(* IEC 61131-3 sources: daoli-st-library/DL_Device (part 15) *)

(* ---- FB_DL_CaseErectFaultSeq.st ---- *)
(*==============================================================================
 * 组件名称 (Component)  : FB_DL_CaseErectFaultSeq
 * 所属子库 (Sublibrary) : DL_Device
 * 当前版本 (Version)    : 1.0.0
 * 兼容性 (Platform)     : CODESYS 3.5+ / TwinCAT 3 / 汇川 InoProShop / 施耐德 Machine Expert
 *                         仅依赖 Standard.library（TON / R_TRIG），零厂商私有库
 * 功能描述 (Function)   : 开箱成型失败重试与吸盘堵塞诊断。bStartCmd 沿启动
 *                         成型吸持：bSuctionCmd 置位等待真空达 fVacOkLevel
 *                         （tonSeek 窗）；达压 → bPickDone 单拍并保持吸持监视
 *                         （中途掉压判 eVacDrop）；超时 → 吹气清理（bBlowOffCmd
 *                         in eRetryPause tRetryPause）后重试，超 nMaxRetry 次
 *                         归因收口：全程真空峰值 <= fVacFloor → eVacClog（吸盘
 *                         堵塞/无真空），曾达压后掉 → eVacDrop，部分真空但
 *                         不足 → eVacTimeout。三成因独立分码（R190 归因唯一）。
 * 来源标签 (Origin)     : ROADMAP 在册空勾 P2（R13 新增行）；判据思想复用既有
 *                         VacuumEjector 件（真空等级判据语义域借鉴），实现与
 *                         码位独立 clean-room，IEC 61131-3 标准语义的道莅防御性实现
 * 边界语义 (Boundary)   : ① 三段 TON 一相一实例（R275）：tonSeek/tonPause/
 *                         tonDrop 各自独立，禁跨相复用；
 *                         ② 归因锁存：故障相按锁存回放，不按当下真空重推断（R28）；
 *                         ③ 重试计数只在收口沿或复位沿清（bStop 中止保留计数，
 *                         作用域在此声明——中止视为本轮未完，重试额度保留）；
 *                         ④ 组态闸：真空等级/地板值/时间/次数全引脚覆盖（R151）。
 * 输出语义 (Fallback)   : 【R191】bEnable = FALSE → 全输出强制 FALSE（吸持是
 *                         执行器指令，失能必须收敛）；eFault 相 → bSuctionCmd
 *                         强制 FALSE（故障先断气源），bError = TRUE。
 * 码位     (Codes)      : 按 R297 范式零 16# 码位硬编码；错误出口 BOOL+ENUM(eCause)，
 *                         码位待主控收口统一派号。
 * 红线自检 (Redline)    : 7 项红线已自检：R1 零全局 ✓｜R2 零物理地址 ✓｜R3 纯 IEC ✓
 *                         R4 组态闸全引脚/容差比较 ✓｜R5 双语同行注释 ✓
 *                         R6 CASE 带 ELSE 兜底迁 eFault ✓
 *                         R7 三 TON + 两 R_TRIG 段 0 无条件刷新，各实例单用途 ✓
 * 验收向量 (Acceptance) : V1 首次达压 → bPickDone 单拍 TRUE，nRetryCnt=0；
 *                         V2 达压后掉压 → eFault，eCause=eVacDrop；
 *                         V3 三次超时且真空峰值恒为地板值 → eCause=eVacClog；
 *                         V4 三次超时峰值 0.5·fVacOkLevel → eCause=eVacTimeout；
 *                         V5 重试期 bBlowOffCmd 电平 TRUE（暂停相内）。
 * 修订历史 (Revision)   : 2026-11-20  v1.0.0  R49 首版（批 2 · 序号 10）
 *==============================================================================*)
TYPE E_DL_CefState :
(
    eIdle       := 0,                        (* 待启动 / Idle *)
    eErect      := 10,                       (* 吸持建立中（真空达压窗） / Erecting, vacuum seek *)
    eHold       := 20,                       (* 吸持保持监视（掉压判据） / Holding, drop watch *)
    eRetryPause := 30,                       (* 吹气清理暂停（重试间隔） / Blow-off pause *)
    eFault      := 90                        (* 故障锁存相 / Fault latched phase *)
);
END_TYPE

TYPE E_DL_CefCause :
(
    eNone        := 0,                       (* 无故障成因 / No cause *)
    eVacClog     := 1,                       (* 吸盘堵塞：全程真空不高于地板值 / Suction clog: vacuum never above floor *)
    eVacDrop     := 2,                       (* 中途掉压：曾达压后失压 / Vacuum drop after reaching level *)
    eVacTimeout  := 3,                       (* 达压超时：部分真空但始终不足 / Vacuum seek timeout, partial only *)
    eCfgIllegal  := 4,                       (* 组态非法 / Illegal config *)
    ePhaseBad    := 5                        (* 非法相位兜底 / Illegal phase fallback *)
);
END_TYPE

FUNCTION_BLOCK FB_DL_CaseErectFaultSeq
VAR_INPUT
    bVacOkLvl   : BOOL := FALSE;             (* 真空达压电平（真空开关或比较器输出直连）[-] / Vacuum-ok level input *)
    fVacReading : LREAL := 0.0;              (* 真空读数（归因诊断用）[kPa] / Vacuum reading for diagnosis *)
    fVacOkLevel : LREAL := 60.0;             (* 达压等级阈值，域 > 0.0 [kPa] / Vacuum ok threshold *)
    fVacFloor   : LREAL := 5.0;              (* 地板值：峰值不高于此判堵塞，域 >= 0.0 且 < fVacOkLevel [kPa] / Vacuum floor for clog verdict *)
    tVacSeek    : TIME := T#3S;              (* 达压窗保持时长，域 > T#0S [ms] / Vacuum seek window *)
    tRetryPause : TIME := T#1S;              (* 吹气清理暂停保持时长，域 > T#0S [ms] / Retry pause hold *)
    nMaxRetry   : INT := 3;                  (* 最大重试次数，域 0..20 [次] / Max retry count *)
    bStartCmd   : BOOL := FALSE;             (* 成型启动命令，上升沿发起 / Start command edge *)
    bStop       : BOOL := FALSE;              (* 中止命令，电平 TRUE 立即断吸回 eIdle（保留重试计数，见边界③） / Stop level, keeps retry count *)
    bEnable     : BOOL := TRUE;              (* 使能，FALSE 全输出强制收敛 [-] / Enable *)
    bReset      : BOOL := FALSE;              (* 复位命令，上升沿清故障锁存与全部状态 [-] / Reset command *)
END_VAR
VAR_OUTPUT
    bSuctionCmd : BOOL;                      (* 吸盘吸持命令输出 [-] / Suction command output *)
    bBlowOffCmd : BOOL;                      (* 吹气清理命令输出（重试暂停相电平）[-] / Blow-off command output *)
    bPickDone   : BOOL;                      (* 本轮吸持达压完成单拍位 [-] / Pick-done single-scan pulse *)
    nRetryCnt   : INT;                       (* 本轮已用重试次数 [次] / Retry count this round *)
    nAttemptCnt : INT;                       (* 本轮尝试总次数（含首次）[次] / Attempt count this round *)
    eState      : E_DL_CefState;             (* 状态出口 / State outlet *)
    eCause      : E_DL_CefCause;             (* 故障成因出口（R190 三成因独立分码） / Fault cause outlet *)
    bError      : BOOL;                       (* 故障锁存标志 [-] / Fault latch flag *)
END_VAR
VAR
    _eState   : E_DL_CefState := E_DL_CefState.eIdle;     (* 内部相位（CASE 唯一写入目标） / Internal phase *)
    _eCause   : E_DL_CefCause := E_DL_CefCause.eNone;     (* 故障成因锁存量 / Latched cause *)
    tonSeek   : TON;                         (* 达压窗计时（eErect 相专用），段 0 无条件调用 / Seek timer, phase-specific *)
    tonPause  : TON;                         (* 吹气暂停计时（eRetryPause 相专用），段 0 无条件调用 / Pause timer, phase-specific *)
    tonDrop   : TON;                         (* 掉压确认计时（eHold 相专用），段 0 无条件调用 / Drop confirm timer, phase-specific *)
    rtStart   : R_TRIG;                      (* 启动沿实例，段 0 无条件调用 / Start edge instance *)
    rtReset   : R_TRIG;                      (* 复位沿实例，段 0 无条件调用 / Reset edge instance *)
    _nRetry   : INT;                         (* 重试计数锁存 [次] / Retry count latch *)
    _nAttempt : INT;                         (* 尝试计数锁存 [次] / Attempt count latch *)
    _fVacMax  : LREAL;                       (* 本轮真空峰值锁存（归因判据源）[kPa] / Vacuum peak latch *)
    _bReached : BOOL;                        (* 本轮曾达压位（掉压归因判据）[-] / Reached-ok latch this round *)
    _bFault   : BOOL;                        (* 故障锁存位 / Latched fault bit *)
    _bCfgBad  : BOOL;                        (* 组态非法当拍量 / Illegal config this scan *)
END_VAR

(* —— 段 0：当拍判据派生 + 实例无条件刷新（R228A，三 TON 各自独立 IN 派生） —— *)
_bCfgBad := (fVacOkLevel <= 0.0) OR (fVacFloor < 0.0) OR (fVacFloor >= fVacOkLevel)   (* 组态闸：等级/地板域及序关系（R151 全引脚覆盖） / Config gate *)
            OR (tVacSeek <= T#0S) OR (tRetryPause <= T#0S) OR (nMaxRetry < 0) OR (nMaxRetry > 20);
rtStart(CLK := bStartCmd);                   (* 启动沿每拍必调 / Start edge every scan *)
rtReset(CLK := bReset);                      (* 复位沿每拍必调 / Reset edge every scan *)
tonSeek(IN := _eState = E_DL_CefState.eErect, PT := tVacSeek);        (* 达压窗随相位派生 / Seek timer phase-derived *)
tonPause(IN := _eState = E_DL_CefState.eRetryPause, PT := tRetryPause);   (* 暂停计时随相位派生 / Pause timer phase-derived *)
tonDrop(IN := _eState = E_DL_CefState.eHold AND NOT bVacOkLvl, PT := tRetryPause);   (* 掉压确认随相位派生（PT 复用暂停时长作为失压容忍窗，语义声明） / Drop confirm timer *)

(* —— 段 1：单拍量预清零（R107） —— *)
bPickDone := FALSE;                          (* 达压完成单拍位预清，唯一分支置位 / Pick pulse preset *)

(* —— 段 2：复位沿处理（作用域：清故障 + 清成因 + 清计数 + 清峰值 + 迁 eIdle，R283 逐项声明） —— *)
IF rtReset.Q THEN
    _bFault := FALSE;                        (* 清故障锁存 / Clear fault *)
    _eCause := E_DL_CefCause.eNone;          (* 清成因 / Clear cause *)
    _nRetry := 0;                            (* 清重试计数 / Clear retry count *)
    _nAttempt := 0;                          (* 清尝试计数 / Clear attempt count *)
    _fVacMax := 0.0;                         (* 清真空峰值 / Clear vacuum peak *)
    _bReached := FALSE;                      (* 清曾达压位 / Clear reached latch *)
    _eState := E_DL_CefState.eIdle;          (* 迁待启动相 / Back to idle *)
END_IF

(* —— 段 3：组态闸故障锁存（R45 配对；锁存至复位沿，R189） —— *)
IF _bCfgBad AND NOT _bFault THEN
    _bFault := TRUE;                         (* 锁存故障位 / Latch fault *)
    _eCause := E_DL_CefCause.eCfgIllegal;    (* 成因：组态非法 / Cause: illegal config *)
    _eState := E_DL_CefState.eFault;         (* 同步迁故障相 / Migrate to fault *)
END_IF

(* —— 段 4：CASE 主状态机（ELSE 兜底迁 eFault，红线 6） —— *)
CASE _eState OF
    E_DL_CefState.eIdle:                     (* 待启动相 / Idle *)
        IF rtStart.Q AND bEnable AND NOT _bFault THEN
            _nAttempt := _nAttempt + 1;      (* 尝试计数递增 / Attempt count advance *)
            _fVacMax := 0.0;                 (* 本轮峰值清零 / Clear round peak *)
            _bReached := FALSE;              (* 本轮曾达压清零 / Clear reached latch *)
            _eState := E_DL_CefState.eErect; (* 进入吸持建立 / Enter erect *)
        END_IF
    E_DL_CefState.eErect:                    (* 吸持建立相 / Erect *)
        IF NOT bEnable OR bStop THEN         (* 失能/中止：断吸回待机（重试计数保留，边界③声明） / Disable or stop *)
            _eState := E_DL_CefState.eIdle;  (* 回待机 / Back to idle *)
        ELSIF bVacOkLvl THEN
            _bReached := TRUE;               (* 曾达压置位 / Reached latch *)
            bPickDone := TRUE;               (* 达压完成单拍脉冲 / Pick-done pulse *)
            _eState := E_DL_CefState.eHold;  (* 进入保持监视 / Enter hold *)
        ELSE
            IF fVacReading > _fVacMax THEN
                _fVacMax := fVacReading;     (* 真空峰值跟踪（NaN 参与比较恒 FALSE，不污染峰值） / Vacuum peak tracking, NaN-safe *)
            END_IF
            IF tonSeek.Q THEN
                _nRetry := _nRetry + 1;      (* 超时计一次重试 / Retry count advance *)
                IF _nRetry > nMaxRetry THEN
                    IF _bReached THEN
                        _eCause := E_DL_CefCause.eVacDrop;      (* 曾达压后失压归因（独立分码，R190） / Drop cause *)
                    ELSIF _fVacMax <= fVacFloor THEN
                        _eCause := E_DL_CefCause.eVacClog;      (* 峰值不高于地板：吸盘堵塞归因 / Clog cause *)
                    ELSE
                        _eCause := E_DL_CefCause.eVacTimeout;   (* 部分真空但不足：超时归因 / Timeout cause *)
                    END_IF
                    _bFault := TRUE;         (* 重试耗尽故障锁存（R45 配对） / Retry exhausted fault *)
                    _eState := E_DL_CefState.eFault;   (* 同步迁故障相 / Migrate to fault *)
                ELSE
                    _eState := E_DL_CefState.eRetryPause;   (* 未耗尽：吹气清理后重试 / Enter retry pause *)
                END_IF
            END_IF
        END_IF
    E_DL_CefState.eHold:                     (* 吸持保持相 / Hold *)
        IF NOT bEnable OR bStop THEN
            _eState := E_DL_CefState.eIdle;  (* 失能/中止回待机 / Back to idle *)
        ELSIF bVacOkLvl THEN
            ;                                (* 吸持正常，无动作 / Holding normal *)
        ELSIF tonDrop.Q THEN                 (* 失压持续到容忍窗 / Drop held to tolerance *)
            _eCause := E_DL_CefCause.eVacDrop;   (* 中途掉压归因（独立分码，R190） / Drop cause *)
            _bFault := TRUE;                 (* 故障锁存（R45 配对） / Latch fault *)
            _eState := E_DL_CefState.eFault; (* 同步迁故障相 / Migrate to fault *)
        END_IF
    E_DL_CefState.eRetryPause:               (* 吹气清理暂停相 / Retry pause *)
        IF NOT bEnable OR bStop THEN
            _eState := E_DL_CefState.eIdle;  (* 失能/中止回待机 / Back to idle *)
        ELSIF tonPause.Q THEN
            _nAttempt := _nAttempt + 1;      (* 新尝试计数 / Attempt count advance *)
            _eState := E_DL_CefState.eErect; (* 重新吸持建立 / Re-enter erect *)
        END_IF
    E_DL_CefState.eFault:                    (* 故障相：先断气源，仅复位沿出 / Fault: suction cut *)
        ;                                    (* 锁存回放（R28） / Replay from latch *)
    ELSE                                     (* 非法相位兜底迁安全态 / Illegal phase fallback *)
        _eState := E_DL_CefState.eFault;     (* 迁故障相 / To fault *)
        _bFault := TRUE;                     (* 同步锁存 / Latch *)
        _eCause := E_DL_CefCause.ePhaseBad;  (* 成因：非法相位 / Cause: illegal phase *)
END_CASE

(* —— 段 5：出口映射（双门控：失能收敛 + 故障断气源，R191/R285 全路径赋值） —— *)
IF (NOT bEnable) OR _bFault OR (_eState = E_DL_CefState.eIdle) THEN
    bSuctionCmd := FALSE;                    (* 失能/故障/待机：吸持强制收敛 / Suction forced off *)
    bBlowOffCmd := FALSE;                    (* 吹气强制收敛 / Blow-off forced off *)
ELSIF _eState = E_DL_CefState.eErect OR _eState = E_DL_CefState.eHold THEN
    bSuctionCmd := TRUE;                     (* 建立/保持相：吸持命令电平 / Suction on *)
    bBlowOffCmd := FALSE;                    (* 吹气关闭 / Blow-off off *)
ELSIF _eState = E_DL_CefState.eRetryPause THEN
    bSuctionCmd := FALSE;                    (* 暂停相断吸 / Suction off *)
    bBlowOffCmd := TRUE;                     (* 吹气清理电平 / Blow-off on *)
ELSE
    bSuctionCmd := FALSE;                    (* 兜底收敛 / Fallback off *)
    bBlowOffCmd := FALSE;                    (* 兜底收敛 / Fallback off *)
END_IF
nRetryCnt := _nRetry;                        (* 重试计数镜像 / Retry count mirror *)
nAttemptCnt := _nAttempt;                    (* 尝试计数镜像 / Attempt count mirror *)
bError := _bFault;                           (* 故障标志镜像 / Fault flag mirror *)
eState := _eState;                           (* 状态出口 / State outlet *)
eCause := _eCause;                           (* 成因出口 / Cause outlet *)
END_FUNCTION_BLOCK

(* ---- FB_DL_CaseSealTapeMonitor.st ---- *)
(*
  FB_DL_CaseSealTapeMonitor  —  封箱胶带缺料/断带监视 / Case sealing tape run-out and break monitor
  分类 Category : DL_Device
  码位 Code     : 16#03_2_0A
  版本 Version  : 1.0.0
  溯源 Source   : ISA-18.2 报警管理语义借鉴 · clean-room 实现，仅借分类/参数域/命名，未复制源码
  功能 Function : 1) 张力 + 光电双判据封箱胶带状态监视（复用 FB_DL_SignalDebounce 去抖）；
                  2) 节拍使能时连续 N 拍「无张力 + 光电同态」才判断带（防单拍尖峰）；
                  3) 缺料与断带独立码值（FB33-3 归因唯一），解除需补料确认 + 复位沿。
  边界 Boundary : ① 节拍使能时连续 N 拍无张力 + 光电同态才判断带（防单拍尖峰）；
                  ② 张力传感器无效冻结判定并置码；
                  ③ 缺料（低张力 + 光电无带）与断带（运动中张力突失）独立码值；
                  ④ 报警解除需补料确认 + 复位沿（双条件可达）；
                  ⑤ 输出三行同向：缺料 → 断带 → 去抖状态。
  依赖 Depends  : FB_DL_SignalDebounce × 2（张力低 / 光电无带去抖，每拍无条件调用）

  码表 Error codes（本件子码步进 16#10，避让邻件码位）:
    16#0002_030A 故障级：组态非法（确认拍数 < 1 / 去抖时长 < 0）
    16#0002_031A 故障级：断带（运动中张力突失 + 光电同态确认，锁存需补料 + 复位沿）
    16#0002_032A 信息级：缺料（低张力 + 光电无带，提示级）/ 张力无效判定冻结（不置 bError）
*)

TYPE E_DL_CstPhase :
(
    eIdle  := 0,  // 空闲 / Idle
    eWatch := 10, // 胶带状态监视 / Tape watching
    eBreak := 20, // 断带锁存 / Tape break latched
    eFault := 90  // 组态故障锁定 / Configuration fault locked
);
END_TYPE

FUNCTION_BLOCK FB_DL_CaseSealTapeMonitor
VAR_INPUT
    bEnable       : BOOL;                           // 总使能，FALSE 回空闲 / Master enable
    bCycleEn      : BOOL;                           // 封箱节拍使能（运动中判定窗口）/ Sealing cycle enable
    bReset        : BOOL;                           // 复位，上升沿清组态故障 / Reset, clears fault
    fTensionN     : REAL;                           // 胶带张力 [N] / Tape tension [N]
    bPhotoSensor  : BOOL;                           // 光电传感（TRUE = 有带）/ Photo sensor, TRUE = tape present
    fTensionLoN   : REAL := 2.0;                    // 张力下限 [N]（低于判无张力）/ Tension low limit [N]
    uBreakConfirm : UINT := 5;                      // 断带确认拍数 [拍] / Break confirm scans
    tDebounce     : TIME := T#100MS;                // 信号去抖时长 [ms] / Signal debounce time
    bTapeRefeed   : BOOL;                           // 补料确认（解除条件之一）/ Tape refeed confirmed
    fEps          : REAL := 1.0E-6;                 // 浮点判零容差 [1] / Floating zero tolerance
END_VAR
VAR_OUTPUT
    bTapeMissing  : BOOL;                           // 缺料标志（提示级）/ Tape missing flag, info level
    bTapeBreak    : BOOL;                           // 断带标志（锁存）/ Tape break flag, latched
    bDebouncing   : BOOL;                           // 去抖进行中标志 / Debouncing flag
    bError        : BOOL;                           // 故障标志，与故障级码配对 / Fault flag
    uErrorId      : UDINT;                          // 事件码，0 = 无事件 / Event code
    eStateOut     : E_DL_CstPhase;                  // 状态机当前态，段尾单点映射 / Phase mapped at tail
END_VAR
VAR
    _eState       : E_DL_CstPhase := E_DL_CstPhase.eIdle;  // 内部状态 / Internal state
    fbDebTension  : FB_DL_SignalDebounce;           // 张力低去抖实例（无条件调用）/ Tension-low debounce
    fbDebPhoto    : FB_DL_SignalDebounce;           // 光电无带去抖实例（无条件调用）/ Photo-no-tape debounce
    rtrReset      : R_TRIG;                         // 复位沿 / Reset edge
    bCfgOk        : BOOL;                           // 组态合法标志 / Configuration valid
    bTensionOk    : BOOL;                           // 张力本拍有效 / Tension valid this scan
    bNoTension    : BOOL;                           // 无张力（去抖后）/ No tension, debounced
    bNoPhoto      : BOOL;                           // 光电无带（去抖后）/ No tape by photo, debounced
    bBreakCond    : BOOL;                           // 断带条件（无张力 + 光电同态）/ Break condition
    uBreakCnt     : UINT;                           // 断带确认计数 [拍] / Break confirm counter
    uFault        : UDINT;                          // 锁存故障码 / Latched fault code
    uInfo         : UDINT;                          // 信息级码 / Information code
END_VAR

(* === 段 0 · 实例刷新 === *)
rtrReset(CLK := bReset);                          // 每拍刷新复位沿

(* === 段 1 · 组态闸 === *)
bCfgOk := (uBreakConfirm >= UINT#1)               // 确认拍数下限
          AND (TIME_TO_REAL(tDebounce) >= 0.0)    // 去抖时长非负
          AND (fTensionLoN >= 0.0)                // 张力下限非负域
          AND (fTensionLoN = fTensionLoN);        // NaN 自反
IF NOT bCfgOk THEN
    uFault := 16#0002_030A;                       // 故障级：组态非法
END_IF
IF rtrReset.Q AND bCfgOk THEN
    uFault := 16#0000;                            // 复位沿清组态锁存（解除路径可达）
END_IF
uInfo := 16#0000;                                 // 信息码每拍清零
bTensionOk := (fTensionN = fTensionN) AND (fTensionN >= 0.0) AND (fTensionN < 1.0E30);  // 张力 NaN 自反 + 非负域

(* === 段 2 · 去抖实例（无条件调用）与双判据合成 === *)
fbDebTension(bRawInput := bTensionOk AND (fTensionN < fTensionLoN),   // 原始判据：张力低于下限
             tRiseDelay := tDebounce,             // 上升去抖
             tFallDelay := tDebounce,             // 下降去抖
             bEnable := bEnable AND bCfgOk,       // 使能透传
             bReset := rtrReset.Q);               // 复位沿透传
fbDebPhoto(bRawInput := (NOT bPhotoSensor),       // 原始判据：光电无带
           tRiseDelay := tDebounce,               // 上升去抖
           tFallDelay := tDebounce,               // 下降去抖
           bEnable := bEnable AND bCfgOk,         // 使能透传
           bReset := rtrReset.Q);                 // 复位沿透传
bNoTension := fbDebTension.bStable;               // 无张力（去抖后）
bNoPhoto := fbDebPhoto.bStable;                   // 光电无带（去抖后）
bDebouncing := fbDebTension.bFiltering OR fbDebPhoto.bFiltering;   // 去抖进行中
bBreakCond := bCycleEn AND bTensionOk AND bNoTension AND bNoPhoto;  // 节拍使能 + 无张力 + 光电同态
bTapeMissing := (NOT bCycleEn) AND bTensionOk AND bNoTension AND bNoPhoto;   // 非节拍缺料（提示级）
IF NOT bTensionOk THEN
    uInfo := 16#0002_032A;                        // 信息级：张力无效判定冻结
    uBreakCnt := UINT#0;                          // 无效拍计数归零（禁污染确认）
END_IF

(* === 段 3 · 断带确认计数（连续 N 拍防单拍尖峰）=== *)
IF bBreakCond THEN
    uBreakCnt := uBreakCnt + UINT#1;              // 断带条件确认计数
    IF uBreakCnt >= uBreakConfirm THEN
        uFault := 16#0002_031A;                   // 故障级：断带锁存（需补料 + 复位沿）
    END_IF
ELSE
    uBreakCnt := UINT#0;                          // 条件消失计数归零
END_IF
bTapeBreak := (uFault = 16#0002_031A);            // 断带出口（锁存态映射）

(* === 段 4 · 主状态机（ENUM + CASE，含 ELSE 兜底）=== *)
CASE _eState OF
E_DL_CstPhase.eIdle :
    IF uFault <> 16#0000 THEN
        _eState := E_DL_CstPhase.eFault;          // 故障优先
    ELSIF bEnable AND bCfgOk THEN
        _eState := E_DL_CstPhase.eWatch;          // 进监视相
    END_IF

E_DL_CstPhase.eWatch :
    IF uFault <> 16#0000 THEN
        _eState := E_DL_CstPhase.eBreak;          // 断带锁存转断带相
    ELSIF (NOT bEnable) OR (NOT bCfgOk) THEN
        _eState := E_DL_CstPhase.eIdle;           // 失能回空闲
    END_IF

E_DL_CstPhase.eBreak :
    (* 解除条件：补料确认 + 复位沿（双条件齐备，路径可达） *)
    IF bTapeRefeed AND rtrReset.Q THEN
        uFault := 16#0000;                        // 复位沿清断带锁存
        uBreakCnt := UINT#0;                      // 确认计数复位
        _eState := E_DL_CstPhase.eWatch;          // 回监视相
    END_IF

E_DL_CstPhase.eFault :
    IF uFault = 16#0000 THEN
        _eState := E_DL_CstPhase.eIdle;           // 解锁回空闲
    END_IF

ELSE
    _eState := E_DL_CstPhase.eFault;              // 非法状态拦截
    uFault := 16#0002_030A;                       // 故障级：相 ID 越界复用组态码段
END_CASE

(* === 段 5 · 输出映射（缺料与断带归因唯一：独立码值独立出口）=== *)
IF NOT bTapeBreak THEN
    bTapeMissing := bTapeMissing AND bTensionOk AND bCfgOk;   // 非断带时缺料提示有效
END_IF
bError := (uFault <> 16#0000);                    // 故障标志仅由故障级码置位（R45 配对）
IF bError THEN
    uErrorId := uFault;                           // 故障级优先上报
ELSE
    uErrorId := uInfo;                            // 否则上报信息级码
END_IF
eStateOut := _eState;                             // 输出枚举段尾单点映射（N2 规则）
END_FUNCTION_BLOCK

(* ---- FB_DL_CellFeederVacuum.st ---- *)
(*
  FB_DL_CellFeederVacuum  —  电芯真空上料吸盘（真空窗 + 泄漏率判据 + 掉料重试） / Cell feeder vacuum cup with vacuum window, leakage-rate verdict and drop retry
  分类 Category : DL_Device
  版本 Version  : 1.0.0
  来源 Source   : t1-5-tcopen — 电芯上料吸盘执行器族深化
  溯源 Origin   : 道莅 clean-room 实现；真空窗确认 + 泄漏率判据 + 有限次重试为公开真空吸取工艺逻辑，未复制任何源码行
  功能 Function : 1) 三段顺控：eVac 抽真空（|fVacKpa - fVacTargetKpa| <= fVacTolKpa 达窗）→
                  eLeak 泄漏率测试窗（tLeak 内 fLeakKpaPerS <= fLeakMaxKpaPerS 且 bPartOn 在位）→
                  eDone；2) 掉料重试：泄漏/在位判据失败或 bPartOn 丢失 → eRetry 重抽，
                  重试计数 nRetry 达 nRetryMax 即故障（计数饱和于 nRetryMax）；
                  3) 抽真空超时、测试窗超时各自归因；
                  4) 故障级单码 052D / 信息级 0433 = 吸取确认完成沿。
  接口 Interface: 输入真空度/泄漏率/在位/三个时间量/重试上限；输出状态 + 吸盘指令 + 码
  边界 Boundary : ① 组态闸：fVacTargetKpa <= 0.0、fVacTolKpa <= 0.0、fLeakMaxKpaPerS <= 0.0、
                  tVacTmo/tLeak/tRetry <= T#0S、nRetryMax = 0 → 052D 锁存；
                  ② 真空度/泄漏率非有限（NaN 自反 + Inf 差值自减）→ 052D 锁存，吸盘保持指令撤销；
                  ③ 重试计数为 UINT，递增前先判饱和（不越界）；④ 三 TON + R_TRIG 段 0 无条件调用；
                  ⑤ 故障相迁出唯一路径 = bReset 上升沿（同时清重试计数）；
                  ⑥ 零全局耦合：无 GVL / VAR_EXTERNAL / %I %Q %M 直接地址。
  依赖 Depends  : Standard.library（TON / R_TRIG）
  码表 Error codes（Device 分段见下，故障窗口 052D / 信息窗口 0433）:
    16#0003_052D 故障级：真空上料故障总码（组态非法 / 抽真空超时 / 泄漏率超限且重试耗尽 / 输入非有限），
                 锁存至 bReset 上升沿；归因见 eCause，不新增码位（派单硬约束单码）
    16#0003_0433 信息级：吸取确认完成沿（进 eDone 单拍）
    分段理由：段 0003 故障带 03A0~03FF 于 R42 用尽，启用 05xx 副带续编，避开 0590~0599 判错位段。
  修订历史 Revision :
    2026-11-19  v1.0.0  R43 首版（批次 4 · 序号 17）
*)

TYPE E_DL_CfvState :
(
    eIdle   := 0,     // 未使能：吸盘指令撤销 / Idle, suction withdrawn
    eVac    := 10,    // 抽真空中 / Evacuating
    eLeak   := 20,    // 泄漏率测试窗 / Leakage test window
    eRetry  := 30,    // 掉料重试重抽中 / Retry re-evacuation
    eDone   := 50,    // 吸取完成 / Pick done
    eFault  := 90     // 故障锁存相 / Fault latched phase
);
END_TYPE

TYPE E_DL_CfvCause :
(
    eNone       := 0, // 无故障成因 / No cause
    eCfgIllegal := 1, // 组态非法 / Illegal configuration
    eVacTmo     := 2, // 抽真空超时 / Evacuation timeout
    eLeakHigh   := 3, // 泄漏率超限且重试耗尽 / Leakage high after retries
    eRetryOut   := 4, // 重试次数耗尽 / Retry exhausted
    eNonFinite  := 5  // 输入非有限 / Non-finite input
);
END_TYPE

FUNCTION_BLOCK FB_DL_CellFeederVacuum
VAR_INPUT
    fVacKpa        : REAL := 0.0;      // 吸盘真空度 [kPa]，正压差量纲 / Cup vacuum level
    fVacTargetKpa  : REAL := 60.0;     // 目标真空度 [kPa]，域 > 0 / Target vacuum level
    fVacTolKpa     : REAL := 3.0;      // 真空度容差 [kPa]，域 > 0 / Vacuum tolerance
    fLeakKpaPerS   : REAL := 0.0;      // 实测泄漏率 [kPa/s] / Measured leakage rate
    fLeakMaxKpaPerS: REAL := 0.5;      // 泄漏率上限 [kPa/s]，域 > 0 / Leakage rate limit
    bPartOn        : BOOL := FALSE;    // 料在位检测（电平）[-] / Part-present detection
    tVacTmo        : TIME := T#5S;     // 抽真空超时 [ms]，域 > 0 / Evacuation timeout
    tLeak          : TIME := T#2S;     // 泄漏率测试窗 [ms]，域 > 0 / Leakage test window
    tRetry         : TIME := T#1S;     // 重试泄压间隔 [ms]，域 > 0 / Retry interval
    nRetryMax      : UINT := 3;        // 最大重试次数 [次]，域 > 0 / Maximum retries
    bStart         : BOOL := FALSE;    // 启动命令（电平）[-] / Start command
    bReset         : BOOL := FALSE;    // 复位命令，上升沿清故障与重试计数 [-] / Reset edge
END_VAR
VAR_OUTPUT
    eState         : E_DL_CfvState;    // 状态出口，段 6 单点映射 / State outlet
    eCause         : E_DL_CfvCause;    // 故障成因出口（R190） / Fault cause outlet
    bSuctionCmd    : BOOL;             // 吸盘真空指令 [-] / Suction vacuum command
    bVacOk         : BOOL;             // 真空达窗镜像 [-] / Vacuum reached mirror
    nRetryCount    : UINT;             // 已重试次数 [次] / Retry count
    bCycleDone     : BOOL;             // 吸取完成标志 [-] / Pick done flag
    bError         : BOOL;             // 故障锁存标志 [-] / Fault latch flag
    nErrId         : UDINT;            // 事件码，0 = 无事件 / Event code
END_VAR
VAR
    _eState        : E_DL_CfvState := E_DL_CfvState.eIdle;   // 内部相位（CASE 唯一写入目标） / Internal phase
    _eCause        : E_DL_CfvCause := E_DL_CfvCause.eNone;   // 故障成因锁存（锁存量） / Latched cause
    tonVac         : TON;              // 抽真空超时计时，每周期无条件调用 / Evacuation timer
    tonLeak        : TON;              // 泄漏测试窗计时，每周期无条件调用 / Leakage window timer
    tonRetry       : TON;              // 重试间隔计时，每周期无条件调用 / Retry interval timer
    rtReset        : R_TRIG;           // 复位沿实例，每周期无条件调用 / Reset edge
    _nRetry        : UINT;             // 重试计数保持量（持久） / Retry counter
    _bVacOk        : BOOL;             // 真空达窗当拍量 [-] / Vacuum verdict
    _bLeakOk       : BOOL;             // 泄漏率达标当拍量 [-] / Leakage verdict
    _bNonFin       : BOOL;             // 输入非有限当拍量 [-] / Non-finite input
    _bCfgBad       : BOOL;             // 组态非法当拍量 [-] / Config illegal
    _bFault        : BOOL;             // 故障锁存位（锁存量） / Latched fault bit
    _uFault        : UDINT;            // 故障码锁存（锁存量） / Latched fault code
    _uInfo         : UDINT;            // 信息码，每拍重算 / Transient info code
END_VAR

(* —— 段 0：沿实例与定时器无条件周期刷新 + 当拍量判据 —— *)
_bVacOk := ABS(fVacKpa - fVacTargetKpa) <= fVacTolKpa;                        // 真空容差窗判据 / Vacuum window
_bLeakOk := fLeakKpaPerS <= fLeakMaxKpaPerS;                                  // 泄漏率判据（单侧直比） / Leakage verdict
_bNonFin := (fVacKpa <> fVacKpa) OR (fLeakKpaPerS <> fLeakKpaPerS)
         OR ((fVacKpa - fVacKpa) <> (fVacKpa - fVacKpa))
         OR ((fLeakKpaPerS - fLeakKpaPerS) <> (fLeakKpaPerS - fLeakKpaPerS)); // NaN 自反 + Inf 差值自减 / NaN and Inf
_bCfgBad := (fVacTargetKpa <= 0.0) OR (fVacTolKpa <= 0.0) OR (fLeakMaxKpaPerS <= 0.0)
            OR (tVacTmo <= T#0S) OR (tLeak <= T#0S) OR (tRetry <= T#0S) OR (nRetryMax = 0);   // 组态非法当拍量 / Config illegal
rtReset(CLK := bReset);                                                       // 复位沿，每拍必调 / Reset edge
tonVac(IN := (_eState = E_DL_CfvState.eVac), PT := tVacTmo);                  // 抽真空超时计时 / Evacuation timer
tonLeak(IN := (_eState = E_DL_CfvState.eLeak), PT := tLeak);                  // 泄漏测试窗计时 / Leakage timer
tonRetry(IN := (_eState = E_DL_CfvState.eRetry), PT := tRetry);               // 重试间隔计时 / Retry timer

(* —— 段 1：单拍量预清零（锁存量与重试计数保持量不入清单） —— *)
_uInfo := 16#0000_0000;            // 信息码每拍重算 / Info recomputed
bSuctionCmd := FALSE;              // 吸盘指令缺省撤销 / Suction default withdrawn
bVacOk := FALSE;                   // 真空镜像缺省 FALSE / Vacuum default
bCycleDone := FALSE;               // 完成标志缺省 FALSE / Done default
nErrId := 16#0000_0000;            // 事件码缺省无事件 / Event code default

(* —— 段 2：复位沿 + 组态域闸 —— *)
IF rtReset.Q THEN                              // rtReset.Q = 当拍量 / current scan
    _bFault := FALSE;                          // 清故障锁存位（锁存量） / Clear fault latch
    _uFault := 16#0000_0000;                   // 清故障锁存码（锁存量） / Clear fault code
    _eCause := E_DL_CfvCause.eNone;            // 清成因（锁存量） / Clear cause
    _nRetry := 0;                              // 清重试计数（锁存量） / Clear retry counter
    IF _eState = E_DL_CfvState.eFault THEN
        _eState := E_DL_CfvState.eIdle;        // 故障相迁出：回未使能 / Fault exit to idle
    END_IF
END_IF
IF _bCfgBad THEN                               // 组态域闸 / Config gate
    _uFault := 16#0003_052D;                   // 故障级：真空上料故障总码（05xx 副带） / Device fault code
    _eCause := E_DL_CfvCause.eCfgIllegal;      // 归因：组态非法 / Cause: illegal config
    _bFault := TRUE;                           // 标志与码位配对（R45） / Flag paired with code
END_IF
IF (NOT _bFault) AND _bNonFin THEN             // 非有限锁存 / Non-finite latch
    _uFault := 16#0003_052D;
    _eCause := E_DL_CfvCause.eNonFinite;       // 归因：非有限 / Cause: non-finite
    _bFault := TRUE;
END_IF

(* —— 段 3：超时 / 泄漏超限 / 掉料（判据当拍量） —— *)
IF (NOT _bFault) AND tonVac.Q THEN             // 抽真空超时 / Evacuation timeout
    _uFault := 16#0003_052D;
    _eCause := E_DL_CfvCause.eVacTmo;          // 归因：抽真空超时 / Cause: evac timeout
    _bFault := TRUE;
END_IF
IF (NOT _bFault) AND (_eState = E_DL_CfvState.eLeak) AND tonLeak.Q THEN
    IF (NOT _bLeakOk) OR (NOT bPartOn) THEN    // 泄漏超限或料不在位 / Leak high or part missing
        IF _nRetry >= nRetryMax THEN           // 重试耗尽 → 故障 / Retries exhausted
            _uFault := 16#0003_052D;
            _eCause := E_DL_CfvCause.eRetryOut;   // 归因：重试耗尽 / Cause: retry exhausted
            _bFault := TRUE;
        ELSE
            _eState := E_DL_CfvState.eRetry;   // 未耗尽：进重试相 / Enter retry
        END_IF
    END_IF
END_IF

(* —— 段 4：故障解除式（R240；全当拍量）：rtReset.Q / NOT _bCfgBad / NOT _bNonFin —— *)
IF rtReset.Q AND (NOT _bCfgBad) AND (NOT _bNonFin) THEN
    _bFault := FALSE;                          // 清故障锁存位（锁存量） / Clear fault latch
    _uFault := 16#0000_0000;                   // 清故障锁存码（锁存量） / Clear fault code
    _eCause := E_DL_CfvCause.eNone;            // 清成因（锁存量） / Clear cause
END_IF

(* —— 段 4A：故障锁存相位迁移闸 —— *)
IF _bFault AND (_eState <> E_DL_CfvState.eFault) THEN
    _eState := E_DL_CfvState.eFault;           // 锁存即入故障相 / Latch enters fault phase
END_IF

(* —— 段 5：相位机（CASE 全覆盖 + ELSE 兜底） —— *)
CASE _eState OF

E_DL_CfvState.eIdle:
    IF bStart AND (NOT _bFault) THEN           // 启动条件 / Start gate
        _nRetry := 0;                          // 新循环清重试计数 / Reset retries for new cycle
        _eState := E_DL_CfvState.eVac;         // 进抽真空相 / Enter evacuation
    END_IF

E_DL_CfvState.eVac:
    bSuctionCmd := TRUE;                       // 真空指令置位（相内承载） / Suction command on
    IF _bVacOk THEN                            // 出口 1：真空达窗 / Vacuum reached
        _eState := E_DL_CfvState.eLeak;        // 进泄漏测试窗 / Enter leakage window
    ELSIF NOT bStart THEN                      // 出口 2：撤启动（R98 双出口） / Start released
        _eState := E_DL_CfvState.eIdle;
    END_IF

E_DL_CfvState.eLeak:
    bSuctionCmd := TRUE;                       // 保持真空指令 / Hold suction
    IF tonLeak.Q THEN                          // 测试窗到时 / Window elapsed
        IF _bLeakOk AND bPartOn THEN           // 泄漏达标且料在位 / Leak OK and part present
            _uInfo := 16#0003_0433;            // 信息级：吸取确认完成沿 / Info: pick confirmed
            _eState := E_DL_CfvState.eDone;    // 进完成相 / Enter done
        ELSE
            _eState := E_DL_CfvState.eRetry;   // 否则进重试相（段 3 已裁决耗尽） / Else retry
        END_IF
    ELSIF NOT bStart THEN                      // 撤启动：中止 / Abort
        _eState := E_DL_CfvState.eIdle;
    END_IF

E_DL_CfvState.eRetry:
    IF tonRetry.Q THEN                         // 重试间隔到 / Retry interval elapsed
        IF _nRetry < nRetryMax THEN            // 计数饱和判定后再递增（不越界） / Saturating increment
            _nRetry := _nRetry + 1;
        END_IF
        _eState := E_DL_CfvState.eVac;         // 回抽真空相重抽 / Back to evacuation
    ELSIF NOT bStart THEN                      // 撤启动：中止 / Abort
        _eState := E_DL_CfvState.eIdle;
    END_IF

E_DL_CfvState.eDone:
    bSuctionCmd := TRUE;                       // 完成相保持吸取（搬送中） / Hold suction during transfer
    IF NOT bStart THEN                         // 撤启动：撤销吸取 / Start released withdraws suction
        _eState := E_DL_CfvState.eIdle;
    END_IF

E_DL_CfvState.eFault:
    ;                                          // 故障相：吸盘指令撤销，仅段 4 复位沿可迁出 / Suction off, reset only

ELSE
    _uFault := 16#0003_052D;                   // 故障级：非法相位兜底（归并总码） / Illegal phase fallback
    _eCause := E_DL_CfvCause.eCfgIllegal;      // 归因：相位非法归并组态 / Cause: phase illegal
    _bFault := TRUE;
    _eState := E_DL_CfvState.eFault;           // 强制回故障相 / Force fault phase

END_CASE

(* —— 段 6：出口单点映射（名实同源；故障相吸盘指令撤销） —— *)
IF _bFault THEN
    bSuctionCmd := FALSE;                      // 故障相吸盘指令强制撤销（安全侧） / Suction forced off
    nErrId := _uFault;                         // 故障锁存码回放 / Replay latched code
ELSE
    nErrId := _uInfo;                          // 信息码 / Transient info
END_IF
bVacOk := _bVacOk AND (NOT _bFault);           // 真空达窗镜像 / Vacuum mirror
nRetryCount := _nRetry;                        // 重试计数出口 / Retry count outlet
bCycleDone := (_eState = E_DL_CfvState.eDone); // 完成标志 / Done flag
bError := _bFault;                             // 故障标志同源 / Flag from latch
eState := _eState;                             // 状态出口 / State outlet
eCause := _eCause;                             // 成因出口 / Cause outlet

END_FUNCTION_BLOCK

(* ---- FB_DL_CellVolumeCheck.st ---- *)
(*
  FB_DL_CellVolumeCheck  —  电芯厚度激光测距校验 / Cell thickness laser-range verification
  分类 Category : DL_Device
  码位 Code     : 16#03_2_01
  版本 Version  : 1.0.0
  溯源 Source   : 道莅自研 clean-room，NE43 语义域参照 NAMUR NE43 公开规范
  功能 Function : 1) 激光测距原始值先按 NE43 判有效性（断线/欠量程/超量程），无效值不得参与超差计算；
                  2) 厚度基准（标定常数）为 0 或非正时拒测并置码；
                  3) 超差判定用公差带 + 迟滞，防边界抖动反复分档。
  边界 Boundary : ① 测距原始域先按 NE43 判有效性，无效值不参与超差计算；
                  ② 厚度基准为 0 或未标定时拒测并置码；
                  ③ 超差判定用公差带 + 迟滞（FB_DL_ToleranceWindow），防边界抖动；
                  ④ 输出三行同向：厚度值 → 判定结果 → 拒测标志。
  依赖 Depends  : FB_DL_ToleranceWindow（公差带 + 迟滞判定，每拍无条件调用）；
                  I_DL_AnalogSensor（内联替代：接口无法直接实例化，NE43 判据本件内联实现，仅引用其 E_DL_SignalQuality 枚举）

  码表 Error codes（本件子码步进 16#10，避让邻件码位）:
    16#0002_0301 故障级：厚度基准（标定常数）非正或未标定，拒测
    16#0002_0311 故障级：公差参数非法（公差 <= 0 或迟滞 > 公差/2）
    16#0002_0321 信息级：测距原始值 NE43 域外（欠量程/超量程/断线），本拍不判超差
*)

TYPE E_DL_CvcPhase :
(
    eIdle    := 0,   // 空闲 / Idle
    eRange   := 10,  // 测距有效域判定 / Range validity check
    eJudge   := 20,  // 厚度公差判定 / Thickness tolerance judgment
    eReject  := 30,  // 拒测 / Measurement rejected
    eFault   := 90   // 故障锁定 / Fault locked
);
END_TYPE

FUNCTION_BLOCK FB_DL_CellVolumeCheck
VAR_INPUT
    bEnable      : BOOL;                          // 总使能，FALSE 回空闲 / Master enable
    bSample      : BOOL := TRUE;                  // 采样使能 / Sampling enable
    bReset       : BOOL;                          // 复位，上升沿清故障与拒测 / Reset
    fDistMm      : REAL;                          // 激光测距原始值 [mm]，量程由组态给定 / Raw laser distance [mm]
    fThickRefMm  : REAL := 0.0;                   // 厚度基准（标定常数）[mm]，域 > 0 才有效 / Thickness reference (calibrated) [mm]
    fTolMm       : REAL := 0.05;                  // 厚度公差半带宽 [mm]，域 > 0 / Thickness tolerance half band [mm]
    fHystMm      : REAL := 0.005;                 // 迟滞回差 [mm]，域 0~公差/2 / Hysteresis [mm]
    fRangeLoMm   : REAL := 0.0;                   // 测距量程下限 [mm] / Range low [mm]
    fRangeHiMm   : REAL := 200.0;                 // 测距量程上限 [mm] / Range high [mm]
    fEps         : REAL := 1.0E-6;                // 浮点判零容差 [1] / Floating zero tolerance
END_VAR
VAR_OUTPUT
    fThickMm     : REAL;                          // 实测厚度 [mm]（激光测距换算后的厚度值）/ Measured thickness [mm]
    eQuality     : E_DL_SignalQuality;            // NE43 信号质量分级（引用既有枚举，不重声明）/ NE43 quality grade
    bInTol       : BOOL;                          // 厚度在公差带内 / Thickness within tolerance
    bOverTol     : BOOL;                          // 超差（带迟滞，保持型）/ Out of tolerance, held
    bReject      : BOOL;                          // 拒测标志（保持型）/ Measurement rejected, held
    bError       : BOOL;                          // 故障标志，与故障级码配对 / Fault flag paired with fault codes
    uErrorId     : UDINT;                         // 事件码，0 = 无事件 / Event code, 0 = none
    eStateOut    : E_DL_CvcPhase;                 // 状态机当前态，段尾单点映射 / Phase mapped at tail
END_VAR
VAR
    _eState      : E_DL_CvcPhase := E_DL_CvcPhase.eIdle;  // 内部状态 / Internal state
    rtrReset     : R_TRIG;                        // 复位沿 / Reset edge
    fbTol        : FB_DL_ToleranceWindow;         // 公差带实例（无条件调用）/ Tolerance window instance
    bCfgOk       : BOOL;                          // 公差组态合法 / Tolerance configuration valid
    bRefOk       : BOOL;                          // 厚度基准有效（已标定）/ Reference valid
    bRangeOk     : BOOL;                          // 测距量程有效（NE43 eGood）/ Range valid
    eQualBuf     : E_DL_SignalQuality;            // NE43 质量暂存 / Quality buffer
    fThickBuf    : REAL;                          // 厚度暂存 [mm] / Thickness buffer
    uFault       : UDINT;                         // 锁存故障码 / Latched fault code
    uInfo        : UDINT;                         // 信息级码 / Information code
END_VAR
VAR CONSTANT
    DL_CVC_RMAX  : REAL := 1000.0;                // 测距量程物理域上限 [mm] / Range domain high [mm]
END_VAR

(* === 段 0 · 实例刷新（无条件周期调用）=== *)
rtrReset(CLK := bReset);                          // 每拍刷新复位沿

(* === 段 1 · NE43 判据（内联替代 I_DL_AnalogSensor，仅引用其质量枚举）=== *)
IF (fDistMm <> fDistMm) OR (ABS(fDistMm) >= 1.0E30) THEN
    eQualBuf := E_DL_SignalQuality.eOpenLoop;     // NaN/Inf：按回路开路处理
ELSIF fDistMm < fRangeLoMm - 1.0 THEN
    eQualBuf := E_DL_SignalQuality.eWireBreakLow; // 低于量程 1 mm 以上：低侧断线
ELSIF fDistMm < fRangeLoMm THEN
    eQualBuf := E_DL_SignalQuality.eUnderRange;   // 量程下沿内：欠量程
ELSIF fDistMm > fRangeHiMm + 1.0 THEN
    eQualBuf := E_DL_SignalQuality.eWireBreakHigh;// 高于量程 1 mm 以上：高侧断线
ELSIF fDistMm > fRangeHiMm THEN
    eQualBuf := E_DL_SignalQuality.eOverRange;    // 量程上沿内：超量程
ELSE
    eQualBuf := E_DL_SignalQuality.eGood;         // 有效测量域
END_IF
eQuality := eQualBuf;                             // 质量分级输出（单点写入）
bRangeOk := (eQualBuf = E_DL_SignalQuality.eGood);    // 仅 eGood 参与超差计算

(* === 段 2 · 组态闸：厚度基准与公差参数 === *)
bRefOk := (fThickRefMm > fEps) AND (fThickRefMm < DL_CVC_RMAX)
          AND (fThickRefMm = fThickRefMm);        // 基准非正/未标定 → 拒测
bCfgOk := (fTolMm > fEps) AND (fHystMm >= 0.0) AND (fHystMm <= (fTolMm * 0.5))
          AND (fRangeHiMm > fRangeLoMm) AND (fTolMm = fTolMm);         // 含 NaN 自反
IF NOT bRefOk THEN
    uFault := 16#0002_0301;                       // 故障级：基准非正或未标定
END_IF
IF NOT bCfgOk THEN
    uFault := 16#0002_0311;                       // 故障级：公差参数非法
END_IF
IF rtrReset.Q AND bRefOk AND bCfgOk THEN
    uFault := 16#0000;                            // 复位沿清锁存（复位路径可达）
    bReject := FALSE;                             // 拒测标志同步复位
    bOverTol := FALSE;                            // 超差标志同步复位
END_IF
uInfo := 16#0000;                                 // 信息码每拍清零

(* === 段 3 · 公差带实例（每拍无条件调用，仅有效值参与）=== *)
fbTol(bEnable := bEnable AND bRangeOk AND bRefOk AND bCfgOk,   // 无效值不参与超差计算
      fTarget := fThickRefMm,                     // 目标厚度 = 标定基准
      fActual := fDistMm,                         // 实测测距（本件口径：测距即厚度）
      fTolerance := fTolMm,                       // 公差半带宽
      fHysteresis := fHystMm);                    // 迟滞防抖
IF bRangeOk THEN
    fThickBuf := fDistMm;                         // 有效值：厚度 = 测距
    fThickMm := fThickBuf;                        // 厚度输出
ELSE
    uInfo := 16#0002_0321;                        // 信息级：测距域外，本拍不判超差
END_IF

(* === 段 4 · 主状态机（ENUM + CASE，含 ELSE 兜底）=== *)
CASE _eState OF
E_DL_CvcPhase.eIdle :
    bInTol := FALSE;                              // 空闲无判定
    IF (uFault = 16#0002_0301) OR (uFault = 16#0002_0311) THEN
        _eState := E_DL_CvcPhase.eFault;          // 组态故障优先
    ELSIF bEnable AND bSample THEN
        _eState := E_DL_CvcPhase.eRange;          // 进入域判定相
    END_IF

E_DL_CvcPhase.eRange :
    IF (NOT bRangeOk) OR (NOT bRefOk) THEN
        bReject := TRUE;                          // 无效/未标定：拒测
        _eState := E_DL_CvcPhase.eReject;
    ELSE
        _eState := E_DL_CvcPhase.eJudge;          // 有效：转公差判定
    END_IF

E_DL_CvcPhase.eJudge :
    bInTol := fbTol.bOk;                          // 公差带内判定（含迟滞）
    IF fbTol.bOk THEN
        bOverTol := FALSE;                        // 恢复合格：解除超差（可到达的解除路径）
    ELSE
        bOverTol := TRUE;                         // 置位型：超差（段尾不清零）
    END_IF
    IF (NOT bEnable) OR rtrReset.Q THEN
        _eState := E_DL_CvcPhase.eIdle;           // 失能/复位回空闲
    ELSIF bSample THEN
        _eState := E_DL_CvcPhase.eRange;          // 连续采样
    END_IF

E_DL_CvcPhase.eReject :
    bReject := TRUE;                              // 拒测标志保持
    bInTol := FALSE;                              // 拒测期不给合格结论
    IF bRangeOk AND bRefOk AND bEnable THEN
        bReject := FALSE;                         // 恢复有效：解除拒测
        _eState := E_DL_CvcPhase.eJudge;
    END_IF

E_DL_CvcPhase.eFault :
    bReject := TRUE;                              // 故障态拒测（安全侧）
    bInTol := FALSE;                              // 不给合格结论
    IF uFault = 16#0000 THEN
        _eState := E_DL_CvcPhase.eIdle;           // 解锁回空闲
    END_IF

ELSE
    _eState := E_DL_CvcPhase.eFault;              // 非法状态拦截
    uFault := 16#0002_0311;                       // 故障级：相 ID 越界
    bInTol := FALSE;                              // 安全侧不给合格结论
    bReject := TRUE;                              // 安全侧拒测
END_CASE
IF NOT bEnable THEN
    _eState := E_DL_CvcPhase.eIdle;               // 失能最高优先回空闲
    bInTol := FALSE;                              // 失能不给合格结论
END_IF

(* === 段 5 · 输出映射（三行同向：厚度 → 判定 → 拒测）=== *)
IF NOT bRangeOk THEN
    bInTol := FALSE;                              // 无效值绝不判合格
END_IF
bError := (uFault <> 16#0000);                    // 故障标志仅由故障级码置位（R45 配对）
IF bError THEN
    uErrorId := uFault;                           // 故障级优先上报
ELSE
    uErrorId := uInfo;                            // 否则上报信息级码
END_IF
eStateOut := _eState;                             // 输出枚举段尾单点映射（N2 规则）
END_FUNCTION_BLOCK

(* ---- FB_DL_ChamberGateValve.st ---- *)
//==============================================================================
// 功能块：FB_DL_ChamberGateValve ｜ 中文名称：真空腔体闸阀双位置互锁驱动
// 所属子库：DL_Device ｜ 版本：v1.0.0 ｜ 兼容：CODESYS V3.5+ / TwinCAT 3 / 汇川 InoProShop
// 功能描述：真空腔体闸阀驱动——开/关到位双反馈确认、抽气侧联锁（抽气中
//           禁开）、双反馈/双命令矛盾防御、移动态超时保护；双输出互斥
//           断言（任一拍 NOT(bOpenOut AND bCloseOut)）结构性成立。
// 开源溯源 (Origin)：道莅 clean-room 防御性实现
// 单位表：阀状态[—]／反馈/命令[—]／超时[ms]
// 错误码表：16#0003_017E 信息级（开/关命令同拍，拒绝并执行关优先——安全
//           侧，不置 bError）/ 16#0003_017F 信息级（抽气中收到开命令，
//           拒绝，不置 bError）/ 16#0003_034E 故障级（双到位反馈同拍为
//           TRUE，到位矛盾，输出全断，置 bError）/ 16#0003_034F 故障级
//           （移动态超时无反馈，输出全断，置 bError）/ 16#0003_0350 故障
//           级兜底（状态机落 ELSE，置 bError）
// 状态机：E_DL_GateValveState（eIdle=0 / eOpening=10 / eClosing=20 /
//           eOpened=30 / eClosed=40 / eFault=99；六态，移动语义按方向
//           拆分为 eOpening/eClosing，对应派单摘要中的 eMoving），CASE 含
//           ELSE 兜底，ELSE 置 0350 并回 eFault
// 边界行为：① 双反馈同拍 TRUE → 故障 034E、输出全断（任何命令都不再
//           输出，直至矛盾消失）；② 双命令同拍 TRUE → 拒绝 + 信息 017E
//           （关优先）；③ 抽气中收到开命令 → 拒绝 + 信息 017F；④ 移动态
//           超时无反馈 → 故障 034F + 输出全断；⑤ 双输出互斥由 IF/ELSE
//           单源赋值结构保证，无显式互斥代码路径。
// 依赖纪律：仅 Standard.library；零同层/跨层调用。
// 修订历史：v1.0.0 2026-11-17 首版（R23 派单 · ROADMAP 半导体 P1 §424）
//==============================================================================

(*------------------------------------------------------------------------------
 * 枚举: E_DL_GateValveState（归属本功能块，同文件发布，全库唯一定义）
 * 含义: 闸阀驱动相位，每个成员在 CASE 中有且仅有一个标签。
 *-----------------------------------------------------------------------------*)
TYPE E_DL_GateValveState :
(
    eIdle    := 0,   // 待机：无命令，输出全断 / Idle, no command, outputs off
    eOpening := 10,  // 开启中：开输出有效，等开到位反馈 / Opening, waiting for the open feedback
    eClosing := 20,  // 关闭中：关输出有效，等关到位反馈 / Closing, waiting for the closed feedback
    eOpened  := 30,  // 已开到位：开反馈确认 / Opened, open feedback confirmed
    eClosed  := 40,  // 已关到位：关反馈确认 / Closed, closed feedback confirmed
    eFault   := 99   // 故障：矛盾/超时/非法状态，输出全断 / Fault, contradiction, timeout or illegal state, outputs off
);
END_TYPE

FUNCTION_BLOCK FB_DL_ChamberGateValve
VAR_INPUT
    bOpenCmd       : BOOL;                  // 开阀命令 [—]，电平有效 / Open command, level active
    bCloseCmd      : BOOL;                  // 关阀命令 [—]，电平有效 / Close command, level active
    bOpenedFb      : BOOL;                  // 开到位反馈 [—] / Opened-position feedback
    bClosedFb      : BOOL;                  // 关到位反馈 [—] / Closed-position feedback
    bPumpingActive : BOOL;                  // 抽气进行中 [—]，抽气中禁开（联锁源） / Pumping active, opening forbidden while pumping
    tFbTimeout     : TIME := T#5S;          // 移动态反馈超时 [ms] / Moving-state feedback timeout [ms]
    bReset         : BOOL;                  // 故障复位 [—]，上升沿退出 eFault / Fault reset, rising edge leaves the fault state
END_VAR
VAR_OUTPUT
    bOpenOut       : BOOL;                  // 开阀输出 [—] / Open output
    bCloseOut      : BOOL;                  // 关阀输出 [—] / Close output
    eValveState    : E_DL_GateValveState;   // 阀相位 [—] / Valve phase
    eErr           : UDINT;                 // 错误码，0 = 无错 / Error code, 0 = no error
    bError         : BOOL;                  // 故障级标志，仅故障级错误置位 / Fault-class flag, set only on fault-level codes
    bValid         : BOOL;                  // 输出可用标志 / Outputs usable flag
END_VAR
VAR
    fbMove         : TON;                   // 移动态反馈超时计时，段 6 无条件刷新 [ms] / Moving feedback timeout
    _eState        : E_DL_GateValveState := E_DL_GateValveState.eIdle; // 当前相位 / Current phase
    _bInit         : BOOL := FALSE;         // 首扫标志，初值 FALSE 取非判定 / First-scan flag, tested negated
    _bFbContradict : BOOL;                  // 双反馈矛盾当拍标志 / Both-feedback contradiction flag
    _bIllegal      : BOOL;                  // 非法状态标志 / Illegal state flag
    _bRejectInfo   : UINT;                  // 拒绝信息码暂存（0 = 无） / Staged rejection info code, zero for none
END_VAR
VAR CONSTANT
    DL_GV_CODE_REJ_BOTH : UINT := 1;        // 双命令拒绝标记 [—] / Rejection marker for dual commands
    DL_GV_CODE_REJ_PUMP : UINT := 2;        // 抽气联锁拒绝标记 [—] / Rejection marker for the pumping interlock
END_VAR

(*------------------------------------------------------------------------------
 * 段 1｜每拍预置：双输出先全断（安全侧），单拍标志预清零
 *      Both outputs cleared first, fail-safe, one-shot flags pre-cleared
 *-----------------------------------------------------------------------------*)
bOpenOut  := FALSE;                         // 开阀输出先清（安全侧） / Open output cleared first
bCloseOut := FALSE;                         // 关阀输出先清（安全侧） / Close output cleared first
eErr      := 16#0000_0000;                  // 错误码每拍重算 / Error code recomputed
bError    := FALSE;                         // 故障标志每拍重算 / Fault flag recomputed
bValid    := FALSE;                         // 可用标志每拍重算 / Usable flag recomputed
_bFbContradict := FALSE;                    // 矛盾标志预清零 / Contradiction flag pre-cleared
_bIllegal := FALSE;                         // 非法状态标志预清零 / Illegal flag pre-cleared
_bRejectInfo := 0;                          // 拒绝标记预清零 / Rejection marker pre-cleared

(*------------------------------------------------------------------------------
 * 段 2｜首扫初始化
 *      First-scan initialisation
 *-----------------------------------------------------------------------------*)
IF NOT _bInit THEN
    _eState := E_DL_GateValveState.eIdle;   // 相位待机起步 / Phase starts idle
    _bInit  := TRUE;                        // 首扫只做一次 / The first scan runs once
END_IF

(*------------------------------------------------------------------------------
 * 段 3｜到位矛盾闸：双反馈同拍 TRUE → 故障 034E 输出全断
 *      Contradiction gate: both position feedbacks TRUE at the same scan
 *-----------------------------------------------------------------------------*)
IF bOpenedFb AND bClosedFb THEN
    _bFbContradict := TRUE;                 // 到位矛盾当拍成立 / Contradiction active this scan
    _eState := E_DL_GateValveState.eFault;  // 转故障态 / Go to the fault state
END_IF

(*------------------------------------------------------------------------------
 * 段 4｜命令防御闸：双命令 → 关优先拒绝；抽气中开命令 → 拒绝
 *      Command defense gates: close priority and the pumping interlock
 *-----------------------------------------------------------------------------*)
IF bOpenCmd AND bCloseCmd THEN
    _bRejectInfo := DL_GV_CODE_REJ_BOTH;    // 双命令拒绝标记 / Dual-command rejection marker
ELSIF bOpenCmd AND bPumpingActive THEN
    _bRejectInfo := DL_GV_CODE_REJ_PUMP;    // 抽气联锁拒绝标记 / Pumping interlock rejection marker
END_IF

(*------------------------------------------------------------------------------
 * 段 5｜移动态超时计时无条件刷新（R40：CASE 之外每拍必调）
 *      Moving timeout refreshed unconditionally per R40
 *-----------------------------------------------------------------------------*)
fbMove(IN := (_eState = E_DL_GateValveState.eOpening)
             OR (_eState = E_DL_GateValveState.eClosing), PT := tFbTimeout); // 移动态反馈超时 / Moving feedback timeout

(*------------------------------------------------------------------------------
 * 段 6｜相位机（只做迁移；输出在段 7 按相置位）
 *      Phase machine, transitions only, outputs assigned in segment seven
 *-----------------------------------------------------------------------------*)
IF NOT _bFbContradict THEN                  // 矛盾当拍冻结相位机 / The machine freezes while the contradiction holds
CASE _eState OF

    E_DL_GateValveState.eIdle:             // 待机：合法命令进入移动态
        IF bCloseCmd AND (NOT bOpenCmd) THEN
            _eState := E_DL_GateValveState.eClosing; // 关命令生效 / Close command accepted
        ELSIF bOpenCmd AND (NOT bCloseCmd) AND (NOT bPumpingActive) THEN
            _eState := E_DL_GateValveState.eOpening; // 开命令生效（抽气中不开） / Open command accepted, not while pumping
        END_IF

    E_DL_GateValveState.eOpening:          // 开启中：到位确认或超时
        IF bOpenedFb THEN
            _eState := E_DL_GateValveState.eOpened;  // 开到位 / Opened confirmed
        ELSIF bCloseCmd AND (NOT bOpenCmd) THEN
            _eState := E_DL_GateValveState.eClosing; // 移动中反向，允许（安全侧就近停） / Reverse while moving, allowed
        ELSIF fbMove.Q THEN
            _eState := E_DL_GateValveState.eFault;   // 超时无反馈，故障全断 / Timeout, fault with outputs off
        END_IF

    E_DL_GateValveState.eClosing:          // 关闭中：到位确认或超时
        IF bClosedFb THEN
            _eState := E_DL_GateValveState.eClosed;  // 关到位 / Closed confirmed
        ELSIF bOpenCmd AND (NOT bCloseCmd) AND (NOT bPumpingActive) THEN
            _eState := E_DL_GateValveState.eOpening; // 移动中反向，允许（抽气联锁仍生效） / Reverse while moving, interlock still applied
        ELSIF fbMove.Q THEN
            _eState := E_DL_GateValveState.eFault;   // 超时无反馈，故障全断 / Timeout, fault with outputs off
        END_IF

    E_DL_GateValveState.eOpened:           // 已开：关命令即转关闭
        IF bCloseCmd THEN
            _eState := E_DL_GateValveState.eClosing; // 关命令生效 / Close command accepted
        END_IF

    E_DL_GateValveState.eClosed:           // 已关：开命令须过抽气联锁
        IF bOpenCmd AND (NOT bPumpingActive) THEN
            _eState := E_DL_GateValveState.eOpening; // 开命令生效 / Open command accepted
        END_IF

    E_DL_GateValveState.eFault:            // 故障：矛盾消失且复位沿才回待机
        IF bReset AND (NOT bOpenedFb) AND (NOT bClosedFb) THEN
            _eState := E_DL_GateValveState.eIdle;    // 原因消失回待机 / The cause is gone, back to idle
        END_IF

    ELSE                                   // 非法状态兜底（R21：CASE 必带 ELSE）
        _bIllegal := TRUE;                 // 标记非法状态 / Flag the illegal state
        _eState   := E_DL_GateValveState.eFault; // 回故障态（安全侧全断） / Back to fault, fail-safe
END_CASE
END_IF

(*------------------------------------------------------------------------------
 * 段 7｜输出置位：IF/ELSE 单源赋值，双输出互斥结构性成立
 *      Output assignment, mutual exclusion holds structurally
 *-----------------------------------------------------------------------------*)
CASE _eState OF
    E_DL_GateValveState.eOpening:          // 开启中：只给开输出 / Opening: only the open output
        bOpenOut := TRUE;                  // 开阀输出 / Open output
    E_DL_GateValveState.eClosing:          // 关闭中：只给关输出 / Closing: only the close output
        bCloseOut := TRUE;                 // 关阀输出 / Close output
    ELSE                                   // 其余相输出全断（含故障） / Otherwise all off, including fault
        bOpenOut  := FALSE;                // 开阀输出断 / Open output off
        bCloseOut := FALSE;                // 关阀输出断 / Close output off
END_CASE

IF _bIllegal THEN
    eErr   := 16#0003_0350;                // 故障级：状态机兜底 / Fault: state machine fallback
    bError := TRUE;                        // 置故障标志 / Raise the fault flag
ELSIF _bFbContradict THEN
    eErr   := 16#0003_034E;                // 故障级：双反馈到位矛盾 / Fault: both-feedback contradiction
    bError := TRUE;                        // 置故障标志 / Raise the fault flag
ELSIF (_eState = E_DL_GateValveState.eFault) THEN
    eErr   := 16#0003_034F;                // 故障级：移动态超时无反馈 / Fault: moving timeout without feedback
    bError := TRUE;                        // 置故障标志 / Raise the fault flag
ELSIF _bRejectInfo = DL_GV_CODE_REJ_BOTH THEN
    eErr := 16#0003_017E;                  // 信息级：双命令拒绝，关优先 / Info: dual commands rejected, close priority
ELSIF _bRejectInfo = DL_GV_CODE_REJ_PUMP THEN
    eErr := 16#0003_017F;                  // 信息级：抽气中开命令拒绝 / Info: open command rejected while pumping
END_IF

bValid := NOT bError;                      // 故障级输出不可用 / Outputs unusable on fault
END_FUNCTION_BLOCK

(* ---- FB_DL_CheckweighZeroTrack.st ---- *)
(*==============================================================================
 * 组件名称 (Component)  : FB_DL_CheckweighZeroTrack
 * 所属子库 (Sublibrary) : DL_Device
 * 当前版本 (Version)    : 1.0.0
 * 兼容性 (Platform)     : CODESYS 3.5 / TwinCAT 3 / 汇川 InoProShop（纯标准元素，零方言）
 * 功能描述 (Function)   : 动态称重零点跟踪与温漂补偿。仅在「空载且无冲击且连续静载满
 *                         静载稳定窗」时更新零点，零点取中值滤波后的原始重量；温漂量按
 *                         (温度 − 标定温度) × 温漂系数 求取并作为诊断量与超限判据输出。
 *                         净重 = 原始重量 − 零点。不做称重采样本身、不做动态滤波调参、
 *                         不做多秤头合并。
 *                         设计反证：温漂量只作为诊断量输出、**不**在净重里二次扣减——零点
 *                         跟踪已把当时的原始值吃进零点，二次扣减会让同一次温漂被扣两遍，
 *                         空载净重出现 ±温漂量 的假残差（本例 0.2 g），正好把真故障掩盖。
 * 溯源 (Origin)         : 道莅 clean-room 防御性实现
 * 本文件内含 (Contains) : TYPE E_DL_ZeroTrackState / FUNCTION_BLOCK FB_DL_CheckweighZeroTrack
 * 依赖 (Depends)        : DL_MathData/FB_DL_MedianFilter（只调用，不复制其内核）
 * 红线自检 (Redline)    : 无外部全局变量、无硬件地址直引 ｜ 全变量中英双语同行注释
 *                         零点漂移限判零防除零 ｜ 非有限用自反比较且保持上次补偿值 ｜
 *                         静载窗定时器与沿实例无条件周期刷新 ｜ 枚举显式赋值 ｜ CASE 含 ELSE
 *                         冻结状态量带解除路径（失能一拍解除），无只置不销状态
 * 错误码表 (Codes)      : 16#0003_03A7 就绪（跟踪正常，含零点未更新但无故障）
 *                         16#0003_03A8 故障级 输入/组态非法（温度非有限、漂移限 ≤0、稳定窗
 *                                    出域）。反证句：温度丢值与「真实 0 ℃ 冷库工况」在数值
 *                                    上同为 0，只能靠非有限判据区分，故必须独立成码
 *                         16#0003_03A9 故障级 相对标定累计漂移超限，零点跟踪冻结（继续跟踪
 *                                    会把误差吃进零点）。反证句：超限事实无法由 03AA「窗未
 *                                    满足」观测，故独立成码
 *                         16#0003_03AA 信息级 跟踪窗未满足，零点保持（不置故障级标志）
 *                         16#0003_03AB 预留：本版不发码（下一轮区间起点，禁止回填）
 * 修订历史 (Revision)   : 2026-11-17  v1.0.0  首版入库 · R28 · 阶段三批 1
 * 验收向量 (Acceptance) : 正向 空载原始 200.0 g 连续静载 1 s、温度 20→30 ℃、系数
 *                         0.02 g/K → 漂移 +0.2 g、零点取 200.0 g、净重 0.0 g、跟踪计数 +1
 *                         反向 空载判据为假且放 500 g 砝码 30 s → 零点不动、净重 500 g；
 *                         温度给 NaN → 16#0003_03A8 且漂移量保持上次值；漂移限给 0 →
 *                         16#0003_03A8；漂移 0.2 g 超限 0.1 g → 16#0003_03A9 且跟踪冻结
 *============================================================================*)

(*-----------------------------------------------------------------------------
 * 枚举: E_DL_ZeroTrackState（归属本功能块，同文件发布，全库唯一定义）
 * 含义: 零点跟踪相位，每个成员在 CASE 中有且仅有一个标签。
 *----------------------------------------------------------------------------*)
TYPE E_DL_ZeroTrackState :
(
    eIdle    := 0,    // 未跟踪：窗条件不满足或禁用 / Not tracking, the window condition is unsatisfied or the function is disabled
    eWatching := 10,  // 窗口计时中：静载计时未满 / Watching, the static window is still counting
    eTracked := 20,   // 本窗已落零点：等条件消失后再开新窗 / Zero latched for this window, waiting for the condition to disappear
    eFrozen  := 99    // 冻结：漂移超限，零点禁止更新 / Frozen, the drift limit was exceeded and the zero must not be updated
);
END_TYPE

FUNCTION_BLOCK FB_DL_CheckweighZeroTrack
VAR_INPUT
    bEnable        : BOOL := FALSE;       // 使能 / Enable
    fWeightRaw_g   : REAL := 0.0;         // 原始毛重 [g]，域 ±50000 / Raw gross weight in grammes, domain plus minus 50000
    bBeltEmpty     : BOOL := FALSE;       // 空载判据（皮带无料） / Belt empty criterion
    bShockActive   : BOOL := FALSE;       // 冲击抑制窗有效（本拍禁止跟踪） / Shock suppression window active, tracking forbidden
    tStableWin     : TIME := T#1S;        // 静载稳定窗 [ms]，域 200ms~10s / Static stability window, domain 200 ms to 10 s
    fTemp_C        : REAL := 20.0;        // 传感器温度 [℃]，域 -20~80 / Sensor temperature in degrees Celsius, domain minus 20 to 80
    fTempRef_C     : REAL := 20.0;        // 标定温度 [℃]，域 -20~80 / Calibration temperature in degrees Celsius
    fDriftCoef_gK  : REAL := 0.02;        // 温漂系数 [g/K]，域 ±0.5 / Temperature drift coefficient in grammes per kelvin, domain plus minus 0.5
    fZeroDevMax_g  : REAL := 5.0;         // 零点漂移限 [g]，域 0.1~50 / Zero drift limit in grammes, domain 0.1 to 50
END_VAR
VAR_OUTPUT
    fZeroOut_g     : REAL;                // 当前零点 [g] / Current zero offset in grammes
    fNetOut_g      : REAL;                // 去皮净重 [g] / Net weight after tare in grammes
    bInWindow      : BOOL;                // 处于合法跟踪窗 / Inside the legal tracking window
    uTrackCnt      : UDINT;               // 零点更新次数 [次] / Zero update count
    fDriftTotal_g  : REAL;                // 相对标定累计温漂 [g]（诊断量，不在净重里二次扣减） / Accumulated temperature drift in grammes, diagnostic only
    bError         : BOOL;                // 故障级标志，仅故障级码置位 / Fault-class flag, set on fault codes only
    eErr           : UDINT;               // 错误码，段位 16#0003_xxxx / Error code in segment 16#0003_xxxx
END_VAR
VAR
    _eState        : E_DL_ZeroTrackState := E_DL_ZeroTrackState.eIdle; // 当前相位 / Current phase
    _bInit         : BOOL := FALSE;       // 首扫标志，取非判定 / First-scan flag, tested negated
    _bWindowOk     : BOOL;                // 窗条件成立（空载 + 无冲击 + 使能） / Window condition satisfied
    _bFrozen       : BOOL;                // 漂移超限冻结状态量（冻结门控挂状态，不挂单拍标志） / Drift freeze state quantity, never a one-shot flag
    _bCfgOk        : BOOL;                // 组态合法标志 / Configuration valid flag
    _fZero         : REAL := 0.0;         // 零点内部副本 [g] / Internal zero offset copy
    _fDrift        : REAL := 0.0;         // 漂移内部副本（非有限时保持）[g] / Internal drift copy, held when the input is not finite
    _fSample       : REAL := 0.0;         // 参与跟踪的重量样本 [g] / Weight sample used for tracking
    _tStableWinEff : TIME := T#1S;        // 生效静载窗（域钳制后） / Effective stability window after clamping
    _tonStable     : TON;                 // 静载窗计时 / Static window timer
    _rtrigWin      : R_TRIG;              // 静载窗计时满上升沿 / Rising edge of the window-full signal
    _fbFilter      : FB_DL_MedianFilter;  // 中值滤波委托实例 / Delegated median filter instance
END_VAR
VAR CONSTANT
    DL_ZT_READY     : UDINT := 16#0003_03A7;  // 就绪码 / Ready code
    DL_ZT_INPUT_BAD : UDINT := 16#0003_03A8;  // 故障级输入/组态非法码 / Fault code for a bad input or configuration
    DL_ZT_DRIFT     : UDINT := 16#0003_03A9;  // 故障级漂移超限码 / Fault code for drift overflow
    DL_ZT_WIN_OFF   : UDINT := 16#0003_03AA;  // 信息级窗未满足码 / Info code for an unsatisfied window
    DL_ZT_WIN_LO    : TIME := T#200MS;        // 静载窗下限 / Stability window lower bound
    DL_ZT_WIN_HI    : TIME := T#10S;          // 静载窗上限 / Stability window upper bound
    DL_ZT_DEV_LO    : REAL := 0.1;            // 漂移限下限 [g] / Drift limit lower bound
    DL_ZT_DEV_HI    : REAL := 50.0;           // 漂移限上限 [g] / Drift limit upper bound
    DL_ZT_COEF_HI   : REAL := 0.5;            // 温漂系数绝对值上限 [g/K] / Absolute drift coefficient bound
    DL_ZT_TEMP_LO   : REAL := -20.0;          // 温度下限 [℃] / Temperature lower bound
    DL_ZT_TEMP_HI   : REAL := 80.0;           // 温度上限 [℃] / Temperature upper bound
END_VAR

// 段 1｜输出与单拍标志预置
bError := FALSE;                                    // 故障标志预清 / Fault flag pre-cleared
eErr := 0;                                          // 错误码预清 / Error code pre-cleared
bInWindow := FALSE;                                 // 窗标志预清 / Window flag pre-cleared

// 段 2｜沿检测无条件周期刷新（严禁置于分支内）
_rtrigWin(CLK := _tonStable.Q);                     // 静载窗计时满沿 / Window-full edge

// 段 3｜首扫初始化（判据取非，R19）：首扫以当前原始重量作为零点起点
IF NOT _bInit THEN
    _fZero := fWeightRaw_g;                         // 零点初始取当前原始值 [g] / The zero starts from the present raw value
    fZeroOut_g := _fZero;                           // 零点出口 [g] / Zero output
    _eState := E_DL_ZeroTrackState.eIdle;           // 相位待机起步 / Phase starts idle
    _bInit := TRUE;                                 // 首扫只做一次 / The first scan runs once
END_IF

// 段 3.5｜冻结解除路径（本件无独立复位引脚，约定「失能一拍」为复位路径，防状态量只置不销）
IF NOT bEnable THEN
    _bFrozen := FALSE;                              // 失能即解除冻结，再使能后重新评估漂移 / A disable pulse releases the freeze, the drift is re-evaluated after re-enabling
END_IF

// 段 4｜中值滤波委托（无条件调用；窗口 5 点，禁用拍不出新样本）
_fbFilter(fIn := fWeightRaw_g, bSample := (bEnable AND NOT bShockActive), nWindow := 5, bClear := FALSE);
_fSample := fWeightRaw_g;                           // 缺省样本取原始值 [g] / The default sample is the raw weight
IF _fbFilter.bValid THEN
    _fSample := _fbFilter.fMedian;                  // 滤波有效则取中值 [g] / Use the median when the filter is valid
END_IF

// 段 5｜组态合法性（漂移限判零防除零；稳定窗与系数出域即组态错）
_bCfgOk := NOT ((fZeroDevMax_g <> fZeroDevMax_g) OR ((fZeroDevMax_g - fZeroDevMax_g) <> (fZeroDevMax_g - fZeroDevMax_g)))
        AND (fZeroDevMax_g >= DL_ZT_DEV_LO) AND (fZeroDevMax_g <= DL_ZT_DEV_HI)
        AND (ABS(fDriftCoef_gK) <= DL_ZT_COEF_HI)
        AND (tStableWin >= DL_ZT_WIN_LO) AND (tStableWin <= DL_ZT_WIN_HI)
        AND (fTempRef_C >= DL_ZT_TEMP_LO) AND (fTempRef_C <= DL_ZT_TEMP_HI);
_tStableWinEff := LIMIT(DL_ZT_WIN_LO, tStableWin, DL_ZT_WIN_HI);   // 生效静载窗钳制 [ms] / Effective stability window after clamping

// 段 6｜温漂求取（温度非有限 → 保持上次漂移值 + 故障码，绝不写 0 掩盖故障）
IF (fTemp_C <> fTemp_C) OR ((fTemp_C - fTemp_C) <> (fTemp_C - fTemp_C)) OR (fTemp_C < DL_ZT_TEMP_LO) OR (fTemp_C > DL_ZT_TEMP_HI) THEN
    eErr := DL_ZT_INPUT_BAD;                        // 故障级：温度非有限或出域，漂移值保持上次 / Fault, temperature not finite, drift held
    bError := TRUE;
ELSE
    _fDrift := (fTemp_C - fTempRef_C) * fDriftCoef_gK;  // 相对标定温度的温漂量 [g] / Drift referred to the calibration temperature
END_IF
IF NOT _bCfgOk THEN
    eErr := DL_ZT_INPUT_BAD;                        // 故障级：组态非法 / Fault, bad configuration
    bError := TRUE;
END_IF
fDriftTotal_g := _fDrift;                           // 漂移诊断量出口 [g] / Drift diagnostic output

// 段 7｜漂移超限闸（超限即冻结零点跟踪；冻结门控挂状态量，不挂单拍标志）
IF ABS(_fDrift) > fZeroDevMax_g THEN
    _bFrozen := TRUE;                               // 冻结状态置位（状态量保持） / Freeze state set and held
    _eState := E_DL_ZeroTrackState.eFrozen;         // 相位转冻结 / Phase to frozen
    eErr := DL_ZT_DRIFT;                            // 故障级：累计漂移超限 / Fault, accumulated drift beyond the limit
    bError := TRUE;
END_IF

// 段 8｜静载窗计时无条件刷新（仅窗条件成立时计时）
_bWindowOk := bEnable AND bBeltEmpty AND (NOT bShockActive) AND _bCfgOk
          AND NOT ((fWeightRaw_g <> fWeightRaw_g) OR ((fWeightRaw_g - fWeightRaw_g) <> (fWeightRaw_g - fWeightRaw_g)));
_tonStable(IN := _bWindowOk AND (NOT _bFrozen), PT := _tStableWinEff);
bInWindow := _bWindowOk AND (NOT _bFrozen);         // 合法跟踪窗标志 / Legal tracking window flag

// 段 9｜零点跟踪状态机（ENUM + CASE + ELSE 兜底）
CASE _eState OF

    E_DL_ZeroTrackState.eIdle:                      // 未跟踪：窗条件成立则开窗计时
        IF bInWindow THEN
            _eState := E_DL_ZeroTrackState.eWatching;   // 进入窗口计时 / Enter the window counting phase
        ELSE
            IF bEnable THEN
                eErr := DL_ZT_WIN_OFF;              // 信息级：窗未满足，零点保持 / Info, the window is unsatisfied and the zero is held
            ELSE
                eErr := DL_ZT_READY;                // 禁用为正常停机 / Disable is a normal stop
            END_IF
        END_IF

    E_DL_ZeroTrackState.eWatching:                  // 窗口计时中：计时满即落零点
        IF NOT bInWindow THEN
            _eState := E_DL_ZeroTrackState.eIdle;   // 条件消失：退出本月窗口 / Condition lost, leave the window
            eErr := DL_ZT_WIN_OFF;                  // 信息级：窗未满足，零点保持 / Info, the window is unsatisfied and the zero is held
        ELSIF _rtrigWin.Q THEN
            _fZero := _fSample;                     // 落零点 = 窗内中值 [g] / Latch the zero from the window median
            fZeroOut_g := _fZero;                   // 零点出口 [g] / Zero output
            uTrackCnt := uTrackCnt + 1;             // 跟踪计数 +1 [次] / Tracking count incremented
            _eState := E_DL_ZeroTrackState.eTracked; // 本窗已落点 / Zero latched for this window
            eErr := DL_ZT_READY;                    // 就绪码 / Ready code
        END_IF

    E_DL_ZeroTrackState.eTracked:                   // 本窗已落点：等条件消失后再开新窗（防同窗重复落点）
        IF NOT bInWindow THEN
            _eState := E_DL_ZeroTrackState.eIdle;   // 条件消失：允许下一次跟踪 / Condition lost, the next tracking may start
        END_IF

    E_DL_ZeroTrackState.eFrozen:                    // 冻结：零点禁止更新，漂移回落后由复位路径解除
        IF NOT _bFrozen THEN
            _eState := E_DL_ZeroTrackState.eIdle;   // 冻结已解除（外部复位后） / Freeze released after an external reset
        ELSE
            eErr := DL_ZT_DRIFT;                    // 故障级：冻结保持 / Fault, the freeze is held
            bError := TRUE;
        END_IF

    ELSE
        // 非法状态兜底（故障级，组态非法码承载）
        eErr := DL_ZT_INPUT_BAD;                    // 故障级：非法相位 / Fault, illegal phase
        bError := TRUE;
        _eState := E_DL_ZeroTrackState.eIdle;

END_CASE

// 段 10｜净重与零点出口（净重单点写入；零点在跟踪路径写入，此处保持）
fZeroOut_g := _fZero;                               // 零点出口（单点回放）[g] / Zero output replayed from the internal copy
fNetOut_g := fWeightRaw_g - _fZero;                 // 去皮净重 [g] / Net weight after tare in grammes
END_FUNCTION_BLOCK

(* ---- FB_DL_CipCaneJuiceLineSeq.st ---- *)
(*
  Component : FB_DL_CipCaneJuiceLineSeq
  Category  : DL_Device
  Type      : FB
  Complexity: C2
  VERSION   : v1.0.0
  功能      : 蔗汁线 CIP 五步清洗时序：ENUM 九态（Idle/PreRinse/Caustic/Intermediate/Rinse/Acid/Final/Done/Fault），按步计时推进，漂洗类步按回液电导早退，单步超时联锁。
  开源溯源  : 道莅原创 clean-room 自研（无外部代码引用）｜License: MIT
  边界条件  : ① 六段步时长与单步超时均须非 0、回液电导合格限须 > 1e-9，否则拒启动并锁故障；
              ② 回液电导早退仅对 Intermediate/Rinse/Final 三个漂洗类步生效，酸洗与碱洗步只认计时；
              ③ 碱洗步叠加温度下限联锁；单步超时为最高优先级故障出口，锁存至 bReset 上升沿。
*)

TYPE E_DL_CaneCipPhase :
(
    eIdle         := 0,    (* 空闲：等启动沿 / Idle waiting start edge *)
    ePreRinse     := 10,   (* 预冲洗：第 1 步 / Pre-rinse step 1 *)
    eCaustic      := 20,   (* 碱洗：第 2 步 / Caustic wash step 2 *)
    eIntermediate := 30,   (* 中间冲洗：第 3 步 / Intermediate rinse step 3 *)
    eRinse        := 40,   (* 清水冲洗：第 4 步 / Rinse step 4 *)
    eAcid         := 50,   (* 酸洗：第 5 步 / Acid wash step 5 *)
    eFinal        := 60,   (* 终冲洗：第 6 步 / Final rinse step 6 *)
    eDone         := 70,   (* 完成：待撤销 / Done holding *)
    eFault        := 90    (* 故障：锁存待复位 / Fault latched *)
);
END_TYPE

FUNCTION_BLOCK FB_DL_CipCaneJuiceLineSeq
VAR_INPUT
    bEnable    : BOOL;                  (* 使能电平 [-] Enable level *)
    bReset     : BOOL;                  (* 复位上升沿，清故障锁存 [-] Reset edge *)
    bStart     : BOOL;                  (* 启动上升沿 [-] Start edge *)
    fCondUs    : REAL;                  (* 回液电导率 [μS/cm] Return liquor conductivity *)
    fCondOkUs  : REAL;                  (* 回液电导合格限 [μS/cm] Conductivity pass limit *)
    atStepTime : ARRAY[0..5] OF TIME;   (* 六段步时长 [ms] Step durations *)
    tStepMax   : TIME;                  (* 单步超时上限 [ms] Single step timeout *)
    fTempC     : REAL;                  (* 碱洗液温度 [°C] Caustic solution temperature *)
    fTempMinC  : REAL;                  (* 碱洗温度下限 [°C] Caustic temperature lower limit *)
END_VAR
VAR_OUTPUT
    bPumpCmd : BOOL;              (* CIP 循环泵输出 [-] CIP circulation pump output *)
    bValveCmd: BOOL;              (* CIP 进液阀输出 [-] CIP inlet valve output *)
    nStep    : INT;               (* 当前步号 1~6 [-] Current step number *)
    ePhase   : E_DL_CaneCipPhase;     (* 相位出口，段尾单点映射 [-] Phase outlet *)
    bDone    : BOOL;              (* 清洗完成（锁存） [-] CIP done latched *)
    bError   : BOOL;              (* 故障锁存标志 [-] Fault latch flag *)
    uErrId   : UDINT;             (* 事件码，0 = 无事件 [-] Event code *)
END_VAR
VAR
    rtReset   : R_TRIG;   (* 复位沿实例，每拍无条件刷新 / Reset edge *)
    rtStart   : R_TRIG;   (* 启动沿实例，每拍无条件刷新 / Start edge *)
    tonStep   : TON;      (* 当前步计时（每拍重装 PT） / Current step timer *)
    tonStepMax: TON;      (* 单步超时（专用超时件） / Step timeout *)
    _ePhase   : E_DL_CaneCipPhase := E_DL_CaneCipPhase.eIdle;  (* 内部相位 / Internal phase *)
    _bFault   : BOOL;     (* 故障锁存位（锁存量） / Latched fault bit *)
    _uFault   : UDINT;    (* 故障码锁存（锁存量） / Latched fault code *)
    _bDone    : BOOL;     (* 完成锁存位（锁存量） / Latched done bit *)
    _bCfgBad  : BOOL;     (* 组态非法当拍量 [-] Config illegal flag *)
    _bNonFin  : BOOL;     (* 输入非有限当拍量 [-] Non-finite input flag *)
    nIdx      : INT;      (* 步时长表遍历下标 [-] Step time loop index *)
    nStepIdx  : INT;      (* 当前步在时长表中的下标 [-] Step index in duration table *)
    tStepNow  : TIME;     (* 当前步时长（已判界） [ms] Current step duration after bound check *)
    bActive   : BOOL;     (* 处于清洗步中 [-] In washing step flag *)
END_VAR
VAR CONSTANT
    DL_EPS     : REAL := 1.0E-9;   (* 除零判定容差 [无量纲] Divide-by-zero tolerance *)
    DL_IDX_MAX : INT := 5;         (* 步时长表最高下标 [-] Highest step table index *)
    DL_ZERO    : TIME := T#0S;     (* 零时长常量 [-] Zero duration *)
END_VAR

(* —— 段 0｜每拍量预清零（锁存量 _bFault/_uFault/_bDone 不入清单） —— *)
uErrId := 16#0000_0000;
_bCfgBad := FALSE;
_bNonFin := FALSE;

(* —— 段 1｜当前步下标：相位映射到 0~5，判界后再取步时长（禁越界读） —— *)
nStepIdx := 0;
CASE _ePhase OF
E_DL_CaneCipPhase.ePreRinse:     nStepIdx := 0;
E_DL_CaneCipPhase.eCaustic:      nStepIdx := 1;
E_DL_CaneCipPhase.eIntermediate: nStepIdx := 2;
E_DL_CaneCipPhase.eRinse:        nStepIdx := 3;
E_DL_CaneCipPhase.eAcid:         nStepIdx := 4;
E_DL_CaneCipPhase.eFinal:        nStepIdx := 5;
ELSE
    nStepIdx := 0;                        (* 非清洗相：下标归 0，时长不用 *)
END_CASE
tStepNow := DL_ZERO;
IF (nStepIdx >= 0) AND (nStepIdx <= DL_IDX_MAX) THEN
    tStepNow := atStepTime[nStepIdx];
END_IF

(* —— 段 2｜非有限拦截与组态闸（覆盖六段时长、单步超时、电导限） —— *)
IF (fCondUs <> fCondUs) OR ((fCondUs - fCondUs) <> 0.0)
   OR (fTempC <> fTempC) OR ((fTempC - fTempC) <> 0.0)
   OR (fCondOkUs <> fCondOkUs) OR ((fCondOkUs - fCondOkUs) <> 0.0)
   OR (fTempMinC <> fTempMinC) OR ((fTempMinC - fTempMinC) <> 0.0) THEN
    _bNonFin := TRUE;
END_IF
IF (tStepMax = T#0S) OR (fCondOkUs <= DL_EPS) THEN
    _bCfgBad := TRUE;
END_IF
FOR nIdx := 0 TO 5 DO
    IF (nIdx >= 0) AND (nIdx <= DL_IDX_MAX) THEN
        IF atStepTime[nIdx] = T#0S THEN
            _bCfgBad := TRUE;             (* 任一段步时长为 0 判组态非法 *)
        END_IF
    END_IF
END_FOR

(* —— 段 3｜清洗步判定 + 沿与定时器每拍无条件刷新（使能挂 IN 引脚） —— *)
bActive := (_ePhase = E_DL_CaneCipPhase.ePreRinse) OR (_ePhase = E_DL_CaneCipPhase.eCaustic)
           OR (_ePhase = E_DL_CaneCipPhase.eIntermediate) OR (_ePhase = E_DL_CaneCipPhase.eRinse)
           OR (_ePhase = E_DL_CaneCipPhase.eAcid) OR (_ePhase = E_DL_CaneCipPhase.eFinal);
rtReset  (CLK := bReset);
rtStart  (CLK := bStart);
tonStep  (IN := bActive AND (NOT _bFault), PT := tStepNow);
tonStepMax(IN := bActive AND (NOT _bFault), PT := tStepMax);

(* —— 段 4｜复位沿：一次性清干净，回空闲（唯一解除路径，恒可达） —— *)
IF rtReset.Q THEN
    _bFault := FALSE;
    _uFault := 16#0000_0000;
    _bDone := FALSE;
    _ePhase := E_DL_CaneCipPhase.eIdle;
END_IF

(* —— 段 5｜主状态机：九态全覆盖 + ELSE 兜底 —— *)
CASE _ePhase OF
E_DL_CaneCipPhase.eIdle:
    bPumpCmd := FALSE; bValveCmd := FALSE; nStep := 0;
    IF rtStart.Q AND bEnable AND (NOT _bFault) AND (NOT _bCfgBad) AND (NOT _bNonFin) THEN
        _bDone := FALSE;
        _ePhase := E_DL_CaneCipPhase.ePreRinse;
    ELSIF rtStart.Q AND (_bFault OR _bCfgBad OR _bNonFin) THEN
        _bFault := TRUE;                  (* 带病启动拒绝 / Reject start with bad config *)
        _uFault := 16#0030_0001;
        _ePhase := E_DL_CaneCipPhase.eFault;
    END_IF

E_DL_CaneCipPhase.ePreRinse:
    bPumpCmd := TRUE; bValveCmd := TRUE; nStep := 1;
    IF tonStepMax.Q THEN
        _bFault := TRUE; _uFault := 16#0030_0002;   (* 故障级：第 1 步超时 *)
        _ePhase := E_DL_CaneCipPhase.eFault;
    ELSIF tonStep.Q THEN
        _ePhase := E_DL_CaneCipPhase.eCaustic;          (* 迁出条件 1：步计时到 *)
    ELSIF NOT bEnable THEN
        _ePhase := E_DL_CaneCipPhase.eIdle;             (* 迁出条件 2：使能撤销 *)
    END_IF

E_DL_CaneCipPhase.eCaustic:
    bPumpCmd := TRUE; bValveCmd := TRUE; nStep := 2;
    IF tonStepMax.Q THEN
        _bFault := TRUE; _uFault := 16#0030_0003;   (* 故障级：第 2 步超时 *)
        _ePhase := E_DL_CaneCipPhase.eFault;
    ELSIF fTempC < fTempMinC THEN
        _bFault := TRUE; _uFault := 16#0030_0004;   (* 故障级：碱洗温度不足 *)
        _ePhase := E_DL_CaneCipPhase.eFault;
    ELSIF tonStep.Q THEN
        _ePhase := E_DL_CaneCipPhase.eIntermediate;     (* 迁出条件 1：步计时到 *)
    ELSIF NOT bEnable THEN
        _ePhase := E_DL_CaneCipPhase.eIdle;             (* 迁出条件 2：使能撤销 *)
    END_IF

E_DL_CaneCipPhase.eIntermediate:
    bPumpCmd := TRUE; bValveCmd := TRUE; nStep := 3;
    IF tonStepMax.Q THEN
        _bFault := TRUE; _uFault := 16#0030_0005;   (* 故障级：第 3 步超时 *)
        _ePhase := E_DL_CaneCipPhase.eFault;
    ELSIF tonStep.Q THEN
        _ePhase := E_DL_CaneCipPhase.eRinse;            (* 迁出条件 1：步计时到 *)
    ELSIF fCondUs <= fCondOkUs THEN
        _ePhase := E_DL_CaneCipPhase.eRinse;            (* 迁出条件 2：回液电导早退 *)
    ELSIF NOT bEnable THEN
        _ePhase := E_DL_CaneCipPhase.eIdle;             (* 迁出条件 3：使能撤销 *)
    END_IF

E_DL_CaneCipPhase.eRinse:
    bPumpCmd := TRUE; bValveCmd := TRUE; nStep := 4;
    IF tonStepMax.Q THEN
        _bFault := TRUE; _uFault := 16#0030_0006;   (* 故障级：第 4 步超时 *)
        _ePhase := E_DL_CaneCipPhase.eFault;
    ELSIF tonStep.Q THEN
        _ePhase := E_DL_CaneCipPhase.eAcid;             (* 迁出条件 1：步计时到 *)
    ELSIF fCondUs <= fCondOkUs THEN
        _ePhase := E_DL_CaneCipPhase.eAcid;             (* 迁出条件 2：回液电导早退 *)
    ELSIF NOT bEnable THEN
        _ePhase := E_DL_CaneCipPhase.eIdle;             (* 迁出条件 3：使能撤销 *)
    END_IF

E_DL_CaneCipPhase.eAcid:
    bPumpCmd := TRUE; bValveCmd := TRUE; nStep := 5;
    IF tonStepMax.Q THEN
        _bFault := TRUE; _uFault := 16#0030_0007;   (* 故障级：第 5 步超时 *)
        _ePhase := E_DL_CaneCipPhase.eFault;
    ELSIF tonStep.Q THEN
        _ePhase := E_DL_CaneCipPhase.eFinal;            (* 迁出条件 1：步计时到 *)
    ELSIF NOT bEnable THEN
        _ePhase := E_DL_CaneCipPhase.eIdle;             (* 迁出条件 2：使能撤销 *)
    END_IF

E_DL_CaneCipPhase.eFinal:
    bPumpCmd := TRUE; bValveCmd := TRUE; nStep := 6;
    IF tonStepMax.Q THEN
        _bFault := TRUE; _uFault := 16#0030_0008;   (* 故障级：第 6 步超时 *)
        _ePhase := E_DL_CaneCipPhase.eFault;
    ELSIF tonStep.Q THEN
        _bDone := TRUE;
        _ePhase := E_DL_CaneCipPhase.eDone;             (* 迁出条件 1：末步计时到 *)
    ELSIF fCondUs <= fCondOkUs THEN
        _bDone := TRUE;
        _ePhase := E_DL_CaneCipPhase.eDone;             (* 迁出条件 2：回液电导早退 *)
    ELSIF NOT bEnable THEN
        _ePhase := E_DL_CaneCipPhase.eIdle;             (* 迁出条件 3：使能撤销 *)
    END_IF

E_DL_CaneCipPhase.eDone:
    bPumpCmd := FALSE; bValveCmd := FALSE; nStep := 0;
    IF NOT bStart THEN
        _ePhase := E_DL_CaneCipPhase.eIdle;             (* 启动撤销：回空闲 *)
    END_IF

E_DL_CaneCipPhase.eFault:
    bPumpCmd := FALSE; bValveCmd := FALSE;          (* 故障相：泵与阀全部切除 *)

ELSE
    _bFault := TRUE;                                (* 兜底：非法相位锁存 *)
    _uFault := 16#0030_0009;
    _ePhase := E_DL_CaneCipPhase.eFault;
END_CASE

(* —— 段 6｜出口单点映射 —— *)
ePhase := _ePhase;
bDone := _bDone;
bError := _bFault;
IF _bFault AND (_uFault <> 16#0000_0000) THEN
    uErrId := _uFault;                              (* 故障码锁存回放 / Latched fault replay *)
END_IF
END_FUNCTION_BLOCK

(* ---- FB_DL_CleaningBrushWear.st ---- *)
(*
  FB_DL_CleaningBrushWear  —  清扫机器人刷辊磨损与换刷里程 / Cleaning-robot brush wear and replacement mileage
  分类 Category : DL_Device
  码位 Code     : 16#03_2_1A
  段位说明      : 03_2 段低半字节已满，1x 段续号，19 格由 ElMutingGantry 启用，本件启用 1A 格（R192）
  版本 Version  : 1.0.0
  来源 Source   : t2-6-rockwell-aoi — 三分类诊断结构借 T2-6 AOI 语义（里程类 / 电流类 / 组态类）
  溯源 Origin   : clean-room 实现，未复制任何源码行
                  （判据取「磨损累计」语义：里程累计 + 电流趋势窗双判据，非单件越限）
  功能 Function : 1) 里程类：FB_DL_EventCounter 累计里程脉冲 → 折算里程 fWearMeters，
                  达 fWearDistMaxM 判磨损（bWearDist 锁存）；
                  2) 电流类：FB_DL_SignalStatistics 电流趋势窗（均值口径），窗口均值 / 标称电流
                  比值达 fWearRatioMax 判磨损（bWearCur 锁存）；
                  3) 组态类：参数域非法判组态故障（bCfgFault 锁存）；
                  4) 换刷沿 bBrushReplaced：三件基准全量重置（计数 / 运行时长 / 统计窗），诊断归零；
                  5) 伴随量：FB_DL_RuntimeMeter 刷辊累计运行时长（保养随行台账）。
  边界 Boundary : ① 三分类诊断结构（里程 / 电流 / 组态）各有独立码值，归因唯一，禁共用枚举成员（R190）；
                  ② fMetersPerPulse <= 0 里程折算除零守卫：判组态类故障，折算出口置 0；
                  ③ fCurrentNomA <= 0 电流比值除零守卫：判组态类故障，比值出口置 0；
                  ④ 换刷沿用 R_TRIG 捕获后以单拍电平喂三件的复位/清零引脚（沿消费纪律）；
                  ⑤ 无状态机 CASE 主相（诊断型 FB）：故障经独立锁存位承载，无跨相 TON 复用问题。
  依赖 Depends  : FB_DL_EventCounter / FB_DL_RuntimeMeter / FB_DL_SignalStatistics（实例化，引脚按 registry 实名）
  码表 Error codes（本件格 03_2_1A，子码步进 +0x100）:
    16#0003_011A 信息级：换刷重置完成（基准全量归零）
    16#0003_021A 故障级：组态类故障（里程折算系数 / 标称电流 / 阈值 / 窗长域非法），锁存至复位
    16#0003_031A 故障级：里程类磨损（累计里程达阈值），锁存至复位或换刷沿
    16#0003_041A 故障级：电流类磨损（趋势窗均值/标称比达阈值），锁存至复位或换刷沿
    16#0003_051A 信息级：统计窗未满（电流判据尚未生效，bCurReady = FALSE）

  修订历史 Revision :
    2026-11-19  v1.0.0  R39 首版（批次 3 · 序号 12）
*)

TYPE E_DL_BrushDiag :
(
    eNone    := 0,    // 无诊断结论 / No diagnosis
    eConfig  := 10,   // 组态类 / Configuration class
    eMileage := 20,   // 里程类 / Mileage class
    eCurrent := 30,   // 电流类 / Current class
    eBoth    := 40    // 里程 + 电流双判 / Both mileage and current
);
END_TYPE

FUNCTION_BLOCK FB_DL_CleaningBrushWear
VAR_INPUT
    bBrushRun      : BOOL := FALSE;      // 刷辊运行反馈（电平）[-] / Brush running feedback, level
    bDistPulse     : BOOL := FALSE;      // 里程脉冲（上升沿有效）[-] / Mileage pulse, rising edge
    fMetersPerPulse: REAL := 0.01;       // 每脉冲折算里程 [m/脉冲]，域 > 0 / Meters per pulse, must exceed zero
    fCurrentNomA   : REAL := 2.0;        // 刷辊电机标称电流 [A]，域 > 0 / Nominal motor current
    fMotorCurrentA : REAL := 0.0;        // 刷辊电机实测电流 [A] / Measured motor current
    fWearDistMaxM  : REAL := 50000.0;    // 换刷里程阈值 [m]，域 > 0 / Replacement mileage threshold
    fWearRatioMax  : REAL := 1.3;        // 电流磨损比值阈值 [无量纲]，域 > 1 / Current wear ratio threshold
    nStatWindow    : INT  := 32;         // 电流统计窗长 [个]，2..64（越界钳位）/ Current statistics window length
    bBrushReplaced : BOOL := FALSE;      // 换刷指令沿，上升沿重置三件基准 / Brush replaced, rising edge resets baselines
    uDeltaTimeMs   : UDINT := 10;        // 任务周期注入 [ms]（运行时长折算用）/ Task cycle time for runtime meter
    bReset         : BOOL := FALSE;      // 故障复位，上升沿生效 / Fault reset, rising edge
END_VAR
VAR_OUTPUT
    fWearMeters : REAL;                   // 累计磨损里程 [m] / Accumulated wear mileage
    fCurMeanA   : REAL;                   // 电流趋势窗均值 [A] / Current window mean
    fCurRatio   : REAL;                   // 电流比值 = 窗均值 / 标称 [无量纲] / Current ratio mean over nominal
    uRunMinutes : UDINT;                  // 刷辊累计运行时长 [min] / Brush accumulated runtime
    bCurReady   : BOOL;                   // 电流判据生效（统计窗已满）[-] / Current criterion ready, window full
    bWearDist   : BOOL;                   // 里程类磨损锁存 [-] / Mileage wear latch
    bWearCur    : BOOL;                   // 电流类磨损锁存 [-] / Current wear latch
    bCfgFault   : BOOL;                   // 组态类故障锁存 [-] / Configuration fault latch
    eDiag       : E_DL_BrushDiag;         // 三分类诊断出口 / Three-class diagnosis outlet
    bReplaceReq : BOOL;                   // 换刷请求（任一磨损锁存）[-] / Replacement request, any wear latch
    bError      : BOOL;                   // 故障聚合位（任一故障锁存）[-] / Aggregate fault flag
    uErrorId    : UDINT;                  // 事件码，0 = 无事件（故障级锁存回放）/ Event code
END_VAR
VAR
    fbDist    : FB_DL_EventCounter;       // 里程脉冲计数实例（主体首部无条件刷新）/ Mileage pulse counter instance
    fbRun     : FB_DL_RuntimeMeter;       // 刷辊运行时长实例（主体首部无条件刷新）/ Brush runtime meter instance
    fbCur     : FB_DL_SignalStatistics;   // 电流趋势统计窗实例（主体首部无条件刷新）/ Current statistics window instance
    rtPulse   : R_TRIG;                   // 里程脉冲上升沿 / Mileage pulse rising edge
    rtReplaced: R_TRIG;                   // 换刷指令上升沿 / Brush replaced rising edge
    rtReset   : R_TRIG;                   // 故障复位上升沿 / Fault reset rising edge
    _rWearM   : REAL;                     // 里程折算中间量 [m] / Mileage conversion working value
    _rRatio   : REAL;                     // 电流比值中间量 [无量纲] / Current ratio working value
    _uPulseTh : DINT;                     // 里程阈值换算脉冲数 [个] / Mileage threshold in pulse count
    _bInit    : BOOL := FALSE;            // 首扫标志，初值 FALSE，判据 NOT bInit（R19 范式）/ First-scan flag
    _bFault   : BOOL;                     // 故障锁存位 / Latched fault bit
    _uFault   : UDINT;                    // 故障码锁存寄存 / Latched fault code register
    _uInfo    : UDINT;                    // 信息码，每拍重算 / Info code
    _bCfgBad  : BOOL;                     // 组态非法聚合 / Configuration invalid aggregate
END_VAR
VAR CONSTANT
    DL_CBW_INF_CAP  : REAL := 1.0E15;        // 非有限值筛查幅值上限 / Non-finite screening cap
    DL_CBW_RATIO_MIN: REAL := 1.0001;        // 电流比值阈值下限（须大于 1，防阈值=1 误判） / Ratio threshold lower bound
END_VAR

(* —— 段 0：依赖件与边沿实例无条件周期刷新（R182：调用语句不得置于 IF/CASE 内） —— *)
rtPulse(CLK := bDistPulse);                                 // 里程脉冲沿刷新，每拍必调
rtReplaced(CLK := bBrushReplaced);                          // 换刷沿刷新，每拍必调
rtReset(CLK := bReset);                                     // 复位沿刷新，每拍必调
fbDist(bCntUp := rtPulse.Q,                                 // 里程脉冲计数
       bCntDown := FALSE,                                   // 无递减
       bLoad := FALSE,                                      // 无装载
       nPreset := 0,                                        // 装载值（未用）
       bWrap := FALSE,                                      // 饱和口径
       nCompHigh := _uPulseTh,                              // 高阈值 = 里程阈值换算脉冲数
       nCompLow := 0,                                       // 低阈值（未用）
       bReset := rtReplaced.Q);                             // 换刷沿单拍喂复位（沿消费纪律）
fbRun(bRunning := bBrushRun,                                // 刷辊运行时长累计
      uDeltaTimeMs := uDeltaTimeMs,                         // 任务周期注入
      uMaintIntervalMin := UDINT#0,                         // 保养预警关闭（由上层另行组态）
      bMaintAck := FALSE,                                   // 无保养确认
      bReset := rtReplaced.Q);                              // 换刷沿单拍清零
fbCur(fIn := fMotorCurrentA,                                // 电流趋势窗采样
      bSample := bBrushRun,                                 // 仅运行时采样（停机电流不入窗）
      nWindow := nStatWindow,                               // 窗长（组态透传，内部钳位）
      bClear := rtReplaced.Q);                              // 换刷沿单拍清窗

(* —— 段 1：单拍量预清零（锁存量 _uFault/_bFault/bWearDist/bWearCur/bCfgFault 不入清单，R187①） —— *)
_uInfo := 16#0000_0000;             // 信息码每拍重算
_bCfgBad := FALSE;                  // 组态非法预清零
bReplaceReq := FALSE;               // 换刷请求缺省 FALSE（段 6 单点重写）
uErrorId := 16#0000_0000;           // 事件码缺省无事件

(* —— 段 2：组态域闸（覆盖全部参与判据换算的引脚，R151；含除零守卫） —— *)
IF (fMetersPerPulse <= 0.0) OR (ABS(fMetersPerPulse) > DL_CBW_INF_CAP)
   OR (fCurrentNomA <= 0.0) OR (ABS(fCurrentNomA) > DL_CBW_INF_CAP) THEN
    _bCfgBad := TRUE;               // 折算系数/标称电流非法（除零守卫命中）
END_IF
IF (fMotorCurrentA <> fMotorCurrentA) OR (ABS(fMotorCurrentA) > DL_CBW_INF_CAP) OR ((fMotorCurrentA - fMotorCurrentA) <> 0.0) THEN
    _bCfgBad := TRUE;               // 实测电流非有限
END_IF
IF (fWearDistMaxM <= 0.0) OR (fWearRatioMax < DL_CBW_RATIO_MIN) OR (nStatWindow < 2) OR (nStatWindow > 64) THEN
    _bCfgBad := TRUE;               // 阈值/窗长域非法
END_IF

(* —— 段 3：组态类故障锁存与解除（R228-B：rtReset.Q 为输入引脚恒可达） —— *)
IF _bCfgBad THEN
    bCfgFault := TRUE;              // 组态类锁存（独立归因，禁并入磨损类）
    IF NOT _bFault THEN
        _uFault := 16#0003_021A;    // 故障级：组态类（仅首次进入时写入）
        _bFault := TRUE;
    END_IF
END_IF
IF rtReset.Q THEN
    _bFault := FALSE;               // 清聚合故障位
    _uFault := 16#0000_0000;
    bCfgFault := FALSE;             // 组态类解除（重置后由段 2 复判）
END_IF

(* —— 段 4：首扫基准与里程阈值换算（分母已闸 > 0） —— *)
IF NOT _bInit THEN
    _uPulseTh := REAL_TO_DINT(fWearDistMaxM / fMetersPerPulse);   // 里程阈值换算脉冲数（分母已闸）
    IF _uPulseTh < 1 THEN
        _uPulseTh := 1;             // 换算下限兜底（防阈值过小永不比较）
    END_IF
    _bInit := TRUE;
END_IF
IF (fMetersPerPulse > 0.0) AND (NOT bCfgFault) THEN
    _rWearM := DINT_TO_REAL(fbDist.nCount) * fMetersPerPulse;   // 里程折算（分母已闸；计数域内标准转换）
ELSE
    _rWearM := 0.0;                 // 组态故障：折算出口置 0（防御口径）
END_IF
fWearMeters := _rWearM;             // 里程出口镜像

(* —— 段 5：电流判据换算（分母已闸；窗未满只给信息级） —— *)
fCurMeanA := fbCur.fMean;           // 窗均值出口镜像
bCurReady := fbCur.bStatValid;      // 方差/统计有效口径（n >= 2）作为判据生效标志
IF (fCurrentNomA > 0.0) AND (NOT bCfgFault) THEN
    _rRatio := fCurMeanA / fCurrentNomA;      // 电流比值（分母已闸）
ELSE
    _rRatio := 0.0;                 // 组态故障：比值出口置 0（防御口径）
END_IF
fCurRatio := _rRatio;               // 比值出口镜像
IF bCurReady AND (NOT bCfgFault) THEN
    IF _rWearM >= fWearDistMaxM THEN
        bWearDist := TRUE;          // 里程类磨损锁存
    END_IF
    IF _rRatio >= fWearRatioMax THEN
        bWearCur := TRUE;           // 电流类磨损锁存
    END_IF
ELSE
    _uInfo := 16#0003_051A;         // 信息级：判据未生效（窗未满或组态故障）
END_IF
IF (bWearDist OR bWearCur) AND (NOT _bFault) THEN
    IF bWearDist AND bWearCur THEN
        _uFault := 16#0003_041A;    // 双判同锁：电流类码承载（里程类独立位 bWearDist 仍可观测，归因不混叠）
    ELSIF bWearDist THEN
        _uFault := 16#0003_031A;    // 里程类磨损
    ELSE
        _uFault := 16#0003_041A;    // 电流类磨损
    END_IF
    _bFault := TRUE;
END_IF
IF rtReplaced.Q THEN
    bWearDist := FALSE;             // 换刷沿：里程类解除
    bWearCur := FALSE;              // 换刷沿：电流类解除
    _uInfo := 16#0003_011A;         // 信息级：换刷重置完成
END_IF

(* —— 段 6：诊断聚合出口（名实同源） —— *)
uRunMinutes := fbRun.uRunTotalMin;  // 运行时长出口镜像
IF bCfgFault THEN
    eDiag := E_DL_BrushDiag.eConfig;            // 组态类优先归因
ELSIF bWearDist AND bWearCur THEN
    eDiag := E_DL_BrushDiag.eBoth;              // 双判
ELSIF bWearDist THEN
    eDiag := E_DL_BrushDiag.eMileage;           // 里程类
ELSIF bWearCur THEN
    eDiag := E_DL_BrushDiag.eCurrent;           // 电流类
ELSE
    eDiag := E_DL_BrushDiag.eNone;              // 无结论
END_IF
bReplaceReq := bWearDist OR bWearCur;           // 换刷请求 = 任一磨损锁存
bError := bCfgFault OR bWearDist OR bWearCur;   // 故障聚合位
IF bError THEN
    uErrorId := _uFault;            // 故障锁存码回放
ELSE
    uErrorId := _uInfo;             // 信息码
END_IF

END_FUNCTION_BLOCK
